// TwinCAT 3 PLC project xpp_pulsepicker_motion
// ProgramVersion: 3.1.4026.17
// libraries:
//   LCLS_MotionAbstraction, * (SLAC)
//   LCLS_Tc_DevAbs, * (SLAC - LCLS)
//   LCLS_Tc_MotSync, * (SLAC - LCLS)
//   Tc2_EtherCAT, * (Beckhoff Automation GmbH)
//   Tc2_MC2, * (Beckhoff Automation GmbH)
//   Tc2_Standard, * (Beckhoff Automation GmbH)
//   Tc2_System, * (Beckhoff Automation GmbH)
//   TcUnit, * (www.tcunit.org)
// project tree:
//   DUTs/ E_HomeIndexState.TcDUT, E_HomeCenterState.TcDUT, E_ModeSelector.TcDUT, E_PickerState.TcDUT, E_PPStatus.TcDUT, E_StatusIndicator.TcDUT, E_ValidationStep.TcDUT, ST_SpeedProfile.TcDUT
//   GVLs/ GVL_Axes.TcGVL, GVL_Common.TcGVL
//   POUs/ FB_FastClose.TcPOU, FB_FastOpen.TcPOU, FB_HomeToCenter.TcPOU, FB_SpindleHomeToCenter.TcPOU, FB_MoveToNearestClosed.TcPOU, FB_PPEPS.TcPOU, FB_SpindleTaskMonitoring.TcPOU, FB_TriggerManagerEL1124.TcPOU (excluded from build), FB_TriggerSetpointManager.TcPOU, PRG_S.TcPOU, PRG_XY.TcPOU
//   POUs/Test/ FB_HomeToCenter_Tests.TcPOU, FB_PPEPS_Tests.TcPOU, PRG_TEST.TcPOU
//   / TestTask.TcTTO, XYTask.TcTTO, STask.TcTTO
// real-time tasks:
//   TASK XYTask: cycle T#5ms, priority 14, ADS port 350
//   TASK STask: cycle T#250us, priority 12, ADS port 351
//   TASK TestTask: cycle T#10ms, priority 16, ADS port 352
// motion (NC):
//   TASK NC-Task 1 SAF: cycle T#250us, priority 4, ADS port 501
//   TASK NC-Task 1 SVB: cycle T#1ms, priority 8, ADS port 511
//   AXIS Y_Test (id 5)
//     OtherSettings: AllowMotionCmdToSlave=true
//     encoder EncType=1
//     drive DrvType=5
//       Analog: TorqueSetpointScale=10, ScaleFactorActTorque=0.1
//       TimeComp: TaskDelayCycles=1
//     controller CtrType=1
//       CtrPara: PriorControlFactor=1
//         Observer: BandWidth=20
//   AXIS X_Test (id 4)
//     OtherSettings: AllowMotionCmdToSlave=true
//     encoder EncType=1
//     drive DrvType=5
//       Analog: TorqueSetpointScale=10, ScaleFactorActTorque=0.1
//       TimeComp: TaskDelayCycles=1
//     controller CtrType=1
//       CtrPara: PriorControlFactor=1
//         Observer: BandWidth=20
//   AXIS Axis_HomeToCenter_Test1 (id 6)
//     OtherSettings: AllowMotionCmdToSlave=true
//     encoder EncType=1
//     drive DrvType=5
//       Analog: TorqueSetpointScale=10, ScaleFactorActTorque=0.1
//     controller CtrType=1
//       CtrPara: PriorControlFactor=1
//         Observer: BandWidth=20
//   AXIS Axis_HomeToCenter_Test2 (id 7)
//     OtherSettings: AllowMotionCmdToSlave=true
//     encoder EncType=1
//     drive DrvType=5
//       Analog: TorqueSetpointScale=10, ScaleFactorActTorque=0.1
//     controller CtrType=1
//       CtrPara: PriorControlFactor=1
//         Observer: BandWidth=20
//   AXIS Axis_HomeToCenter_Test3 (id 8)
//     OtherSettings: AllowMotionCmdToSlave=true
//     encoder EncType=1
//     drive DrvType=5
//       Analog: TorqueSetpointScale=10, ScaleFactorActTorque=0.1
//     controller CtrType=1
//       CtrPara: PriorControlFactor=1
//         Observer: BandWidth=20
//   AXIS Axis_HomeToCenter_Test4 (id 9)
//     OtherSettings: AllowMotionCmdToSlave=true
//     encoder EncType=1
//     drive DrvType=5
//       Analog: TorqueSetpointScale=10, ScaleFactorActTorque=0.1
//     controller CtrType=1
//       CtrPara: PriorControlFactor=1
//         Observer: BandWidth=20
//   AXIS Axis_HomeToCenter_Test5 (id 10)
//     OtherSettings: AllowMotionCmdToSlave=true
//     encoder EncType=1
//     drive DrvType=5
//       Analog: TorqueSetpointScale=10, ScaleFactorActTorque=0.1
//     controller CtrType=1
//       CtrPara: PriorControlFactor=1
//         Observer: BandWidth=20
//   AXIS Y (id 3)
//     Dynamic: AccelerationMaximum=200, DecelerationMaximum=200, Acceleration=134.468, Deceleration=134.468, Jerk=488.416
//     Velo: RefSearch=0.6383, RefSync=0.6383, SlowManual=0.25, FastManual=0.35, Fast=63.83, Maximum=63.83
//     PositionAreaControl: Range=0.1
//     TargetPosControl: Range=0.1
//     PEHControl: Time=1
//     OtherSettings: PulseDistancePos=0.1, PulseDistanceNeg=0.1
//     encoder EncType=19
//       EncPara: ScaleFactorNumerator=5, ScaleFactorDenominator=1048576, EncMode=3, MaxCount=#xffffffff
//         TimeComp: TimeCompMode=1, EncDelayCycles=4
//     drive DrvType=16
//       DrvPara: MaxCount=#xffffffff, DriveControlDWord=#x00020100
//         Analog: VeloReferenz=70.213, VeloScale=32, TorqueSetpointScale=10, ScaleFactorActTorque=0.1
//         TimeComp: TaskDelayCycles=1
//     controller CtrType=2
//       CtrPara: PriorControlFactor=1
//         PosDiffControl: Range=0.1
//         PID: PosKp=0
//         Observer: BandWidth=20
//   AXIS X (id 2)
//     Dynamic: AccelerationMaximum=80, DecelerationMaximum=80, Acceleration=57.5064, Deceleration=57.5064, Jerk=743.932
//     Velo: RefSearch=0.45, RefSync=0.25, SlowManual=0.25, FastManual=0.25, Fast=7.056, Maximum=7.056
//     PositionAreaControl: Range=0.1
//     TargetPosControl: Range=0.1
//     PEHControl: Time=1
//     OtherSettings: PulseDistancePos=0.1, PulseDistanceNeg=0.1
//     encoder EncType=19
//       EncPara: ScaleFactorNumerator=0.635, ScaleFactorDenominator=1048576, EncMode=3, MaxCount=#xffffffff
//         TimeComp: TimeCompMode=1, EncDelayCycles=4
//     drive DrvType=16
//       DrvPara: MaxCount=#xffffffff, DriveControlDWord=#x00020100
//         Analog: VeloReferenz=7.7616, VeloScale=32, TorqueSetpointScale=10, ScaleFactorActTorque=0.1
//         TimeComp: TaskDelayCycles=1
//     controller CtrType=1
//       CtrPara: PriorControlFactor=1
//         PosDiffControl: Range=0.1
//         PID: PosKp=0
//         Observer: BandWidth=20
//   AXIS Spindle (id 1)
//     General: UnitName=°
//     Dynamic: AccelerationMaximum=47150500, DecelerationMaximum=47150500, Acceleration=2512000, Deceleration=2512000, Jerk=2673789830.50848
//     Velo: RefSearch=82.10526, RefSync=82.10526, SlowManual=15.5263, FastManual=25.1578, Fast=14210.526, Maximum=4000
//     PositionAreaControl: Range=0.1
//     TargetPosControl: Range=0.1
//     BacklashCompensation: Range=-1.25
//     OtherSettings: AllowMotionCmdToSlave=true, PulseDistancePos=0.1, PulseDistanceNeg=0.1
//     encoder EncType=19
//       EncPara: ScaleFactorNumerator=360, ScaleFactorDenominator=1048576, MaxCount=#xffffffff
//     drive DrvType=16
//       DrvPara: MaxCount=#xffffffff, DriveControlDWord=#x00020100
//         Analog: VeloReferenz=7200, TorqueSetpointScale=10, ScaleFactorActTorque=0.1
//         TimeComp: TaskDelayCycles=1
//     controller CtrType=2
//       CtrPara: PriorControlFactor=1
//         PosDiffControl: Range=3
//         PID: PosKp=0
//         Observer: BandWidth=20
// I/O:
//   DEVICE Device 1 (EtherCAT), AmsNetId 172.21.86.248.2.1
//     Term 1 (EK1200) [EK1200-5000 EtherCAT Power supply (2A E-Bus)]
//       Dongle [EL6070 1Ch. Licensing-Terminal]
//       Spindle [EL7062-0000 2Ch. Stepper motor output stage (48V, 3A)]
//         startup 28688:3 := 08 // DRV Outputs Ch.1 / Modes of operation
//         startup 28688:16 := FF7F // DRV Outputs Ch.1 / Positive torque limit value
//         startup 28688:17 := FF7F // DRV Outputs Ch.1 / Negative torque limit value
//         startup 32784:87 := 64 // DRV Amplifier Settings Ch.1 / Position loop velocity feed forward gain
//         startup 32784:109 := 64000000 // DRV Amplifier Settings Ch.1 / Torque feed forward gain
//         startup 32785:52 := A00F0000 // DRV Motor Settings Ch.1 / Configured motor current
//         startup 32784:19 := 1A00 // DRV Amplifier Settings Ch.1 / Current loop proportional gain
//         startup 32784:18 := 1300 // DRV Amplifier Settings Ch.1 / Current loop integral time
//         startup 32784:21 := 51000000 // DRV Amplifier Settings Ch.1 / Velocity loop proportional gain
//         startup 32784:20 := 96000000 // DRV Amplifier Settings Ch.1 / Velocity loop integral time
//       XY [EL7062-0000 2Ch. Stepper motor output stage (48V, 3A)]
//         startup 28688:3 := 08 // DRV Outputs Ch.1 / Modes of operation
//         startup 28688:16 := FF7F // DRV Outputs Ch.1 / Positive torque limit value
//         startup 28688:17 := FF7F // DRV Outputs Ch.1 / Negative torque limit value
//         startup 32784:87 := 64 // DRV Amplifier Settings Ch.1 / Position loop velocity feed forward gain
//         startup 32784:109 := 64000000 // DRV Amplifier Settings Ch.1 / Torque feed forward gain
//         startup 32785:52 := C4090000 // DRV Motor Settings Ch.1 / Configured motor current
//         startup 32784:19 := 2800 // DRV Amplifier Settings Ch.1 / Current loop proportional gain
//         startup 32784:18 := 1200 // DRV Amplifier Settings Ch.1 / Current loop integral time
//         startup 32784:21 := 2B000000 // DRV Amplifier Settings Ch.1 / Velocity loop proportional gain
//         startup 32784:20 := 96000000 // DRV Amplifier Settings Ch.1 / Velocity loop integral time
//         startup 33042:19 := 0000 // DRV Brake Settings Ch.2 / Emergency application timeout
//         startup 33040:51 := 0A00 // DRV Amplifier Settings Ch.2 / Stand still window
//         startup 28944:3 := 08 // DRV Outputs Ch.2 / Modes of operation
//         startup 28944:16 := FF7F // DRV Outputs Ch.2 / Positive torque limit value
//         startup 28944:17 := FF7F // DRV Outputs Ch.2 / Negative torque limit value
//         startup 33040:87 := 64 // DRV Amplifier Settings Ch.2 / Position loop velocity feed forward gain
//         startup 33040:109 := 64000000 // DRV Amplifier Settings Ch.2 / Torque feed forward gain
//         startup 33041:52 := A00F0000 // DRV Motor Settings Ch.2 / Configured motor current
//         startup 33040:19 := 3000 // DRV Amplifier Settings Ch.2 / Current loop proportional gain
//         startup 33040:18 := 2700 // DRV Amplifier Settings Ch.2 / Current loop integral time
//         startup 33040:21 := 66000000 // DRV Amplifier Settings Ch.2 / Velocity loop proportional gain
//         startup 33040:20 := 96000000 // DRV Amplifier Settings Ch.2 / Velocity loop integral time
//       Term 5 (EL9505) [EL9505 Power supply terminal 5V]
//       Trigger [EL1124 4Ch. Dig. Input 5V, 10µs, Sensor Power]
//       Term 7 (EL9011) [EL9011 End Terminal]
// variable links:
//   (this object) <-> Device 1 (EtherCAT)/Term 1 (EK1200)/XY
//     Drive/Inputs/In/nDataIn1 <-> DRV Following error actual value Channel 2/Following error actual value
//     Drive/Inputs/In/nDataIn1 <-> DRV Following error actual value Channel 1/Following error actual value
//     Drive/Inputs/In/nDataIn3[0] <-> DRV Torque actual value Channel 2/Torque actual value
//     Drive/Inputs/In/nDataIn3[0] <-> DRV Torque actual value Channel 1/Torque actual value
//     Drive/Inputs/In/nDcOutputTime <-> InfoData/DcOutputShift
//     Drive/Inputs/In/nState1 <-> DRV Statusword Channel 2/Statusword
//     Drive/Inputs/In/nState1 <-> DRV Statusword Channel 1/Statusword
//     Drive/Inputs/In/nState2 <-> DRV Statusword Channel 2/Statusword @bit 8
//     Drive/Inputs/In/nState2 <-> DRV Statusword Channel 1/Statusword @bit 8
//     Drive/Inputs/In/nState4 @bit 1 <-> WcState/InputToggle
//     Drive/Inputs/In/nState4 <-> WcState/WcState
//     Drive/Outputs/Out/nCtrl1 <-> DRV Controlword Channel 2/Controlword
//     Drive/Outputs/Out/nCtrl1 <-> DRV Controlword Channel 1/Controlword
//     Drive/Outputs/Out/nCtrl2 <-> DRV Controlword Channel 2/Controlword @bit 8
//     Drive/Outputs/Out/nCtrl2 <-> DRV Controlword Channel 1/Controlword @bit 8
//     Drive/Outputs/Out/nDataOut1 <-> DRV Target position Channel 2/Target position
//     Drive/Outputs/Out/nDataOut1 <-> DRV Target position Channel 1/Target position
//     Enc/Inputs/In/nDataIn1 <-> FB Position Channel 2/Position
//     Enc/Inputs/In/nDataIn1 <-> FB Position Channel 1/Position
//     Enc/Inputs/In/nDcInputTime <-> InfoData/DcInputShift
//     Enc/Inputs/In/nState4 @bit 1 <-> WcState/InputToggle
//     Enc/Inputs/In/nState4 <-> WcState/WcState
//     XYTask Inputs/PRG_XY.fbX.fbEncoderScaling.nRawEncoderUDINT <-> FB Position Channel 1/Position
//     XYTask Inputs/PRG_XY.fbX.fbLimSwStatus.bLimitBwd <-> DI Inputs Channel 1/Input 1
//     XYTask Inputs/PRG_XY.fbX.fbLimSwStatus.bLimitFwd <-> DI Inputs Channel 1/Input 2
//     XYTask Inputs/PRG_XY.fbY.fbEncoderScaling.nRawEncoderUDINT <-> FB Position Channel 2/Position
//     XYTask Inputs/PRG_XY.fbY.fbLimSwStatus.bLimitBwd <-> DI Inputs Channel 2/Input 2
//     XYTask Inputs/PRG_XY.fbY.fbLimSwStatus.bLimitFwd <-> DI Inputs Channel 2/Input 1
//   (this object) <-> Device 1 (EtherCAT)/Term 1 (EK1200)/Spindle
//     Drive/Inputs/In/nDataIn1 <-> DRV Following error actual value Channel 1/Following error actual value
//     Drive/Inputs/In/nDataIn3[0] <-> DRV Torque actual value Channel 1/Torque actual value
//     Drive/Inputs/In/nState1 <-> DRV Statusword Channel 1/Statusword
//     Drive/Inputs/In/nState2 <-> DRV Statusword Channel 1/Statusword @bit 8
//     Drive/Inputs/In/nState4 @bit 1 <-> WcState/InputToggle
//     Drive/Inputs/In/nState4 <-> WcState/WcState
//     Drive/Outputs/Out/nCtrl1 <-> DRV Controlword Channel 1/Controlword
//     Drive/Outputs/Out/nCtrl2 <-> DRV Controlword Channel 1/Controlword @bit 8
//     Drive/Outputs/Out/nDataOut1 <-> DRV Target position Channel 1/Target position
//     Enc/Inputs/In/nDataIn1 <-> FB Position Channel 1/Position
//     Enc/Inputs/In/nDataIn3 <-> FB Touch probe 1 pos position Channel 1/TP1 Pos position
//     Enc/Inputs/In/nDataIn5 <-> FB Touch probe 2 pos position Channel 1/TP2 Pos position
//     Enc/Inputs/In/nState4 @bit 1 <-> WcState/InputToggle
//     Enc/Inputs/In/nState4 <-> WcState/WcState
//     Enc/Inputs/In/nState5 <-> FB Touch probe status Channel 1/Touch probe status/TP1 Enable
//     Enc/Inputs/In/nState6 <-> FB Touch probe status Channel 1/Touch probe status/TP2 Enable
//     Enc/Inputs/In/nState5 @bit 7 <-> FB Touch probe status Channel 1/Touch probe status/TP1 Input
//     Enc/Inputs/In/nState6 @bit 7 <-> FB Touch probe status Channel 1/Touch probe status/TP2 Input
//     Enc/Inputs/In/nState5 @bit 2 <-> FB Touch probe status Channel 1/Touch probe status/TP1 Neg value stored
//     Enc/Inputs/In/nState6 @bit 2 <-> FB Touch probe status Channel 1/Touch probe status/TP2 Neg value stored
//     Enc/Inputs/In/nState5 @bit 1 <-> FB Touch probe status Channel 1/Touch probe status/TP1 Pos value stored
//     Enc/Inputs/In/nState6 @bit 1 <-> FB Touch probe status Channel 1/Touch probe status/TP2 Pos value stored
//     Enc/Outputs/Out/nCtrl5 @bit 1 <-> FB Touch probe control Channel 1/Touch probe function/TP1 Continous
//     Enc/Outputs/Out/nCtrl6 @bit 1 <-> FB Touch probe control Channel 1/Touch probe function/TP2 Continous
//     Enc/Outputs/Out/nCtrl5 <-> FB Touch probe control Channel 1/Touch probe function/TP1 Enable
//     Enc/Outputs/Out/nCtrl6 <-> FB Touch probe control Channel 1/Touch probe function/TP2 Enable
//     Enc/Outputs/Out/nCtrl5 @bit 5 <-> FB Touch probe control Channel 1/Touch probe function/TP1 Enable neg edge
//     Enc/Outputs/Out/nCtrl6 @bit 5 <-> FB Touch probe control Channel 1/Touch probe function/TP2 Enable neg edge
//     Enc/Outputs/Out/nCtrl5 @bit 4 <-> FB Touch probe control Channel 1/Touch probe function/TP1 Enable pos edge
//     Enc/Outputs/Out/nCtrl6 @bit 4 <-> FB Touch probe control Channel 1/Touch probe function/TP2 Enable pos edge
//     Enc/Outputs/Out/nCtrl5 @bit 2 <-> FB Touch probe control Channel 1/Touch probe function/TP1 Trigger mode
//     Enc/Outputs/Out/nCtrl6 @bit 2 <-> FB Touch probe control Channel 1/Touch probe function/TP2 Trigger mode
//     STask Inputs/PRG_S.fbHomeIdx.bHomeIndex <-> DI Inputs Channel 1/Encoder C
//     STask Inputs/PRG_S.fbS.fbEncoderScaling.nRawEncoderUDINT <-> FB Position Channel 1/Position
//   (this object) <-> Device 1 (EtherCAT)/Term 1 (EK1200)/Trigger
//     STask Inputs/PRG_S.fbTrigMgr.fbTrigSrc.bTrigger <-> Channel 1/Input
//   (this object) <-> NC-Task 1 SAF/Axes/Axis_HomeToCenter_Test1
//     TestTask Inputs/PRG_TEST.fb_HomeToCenter_Tests.fbAxisRef[1].NcToPlc <-> Outputs/ToPlc
//     TestTask Outputs/PRG_TEST.fb_HomeToCenter_Tests.fbAxisRef[1].PlcToNc <-> Inputs/FromPlc
//   (this object) <-> NC-Task 1 SAF/Axes/Axis_HomeToCenter_Test2
//     TestTask Inputs/PRG_TEST.fb_HomeToCenter_Tests.fbAxisRef[2].NcToPlc <-> Outputs/ToPlc
//     TestTask Outputs/PRG_TEST.fb_HomeToCenter_Tests.fbAxisRef[2].PlcToNc <-> Inputs/FromPlc
//   (this object) <-> NC-Task 1 SAF/Axes/Axis_HomeToCenter_Test3
//     TestTask Inputs/PRG_TEST.fb_HomeToCenter_Tests.fbAxisRef[3].NcToPlc <-> Outputs/ToPlc
//     TestTask Outputs/PRG_TEST.fb_HomeToCenter_Tests.fbAxisRef[3].PlcToNc <-> Inputs/FromPlc
//   (this object) <-> NC-Task 1 SAF/Axes/Axis_HomeToCenter_Test4
//     TestTask Inputs/PRG_TEST.fb_HomeToCenter_Tests.fbAxisRef[4].NcToPlc <-> Outputs/ToPlc
//     TestTask Outputs/PRG_TEST.fb_HomeToCenter_Tests.fbAxisRef[4].PlcToNc <-> Inputs/FromPlc
//   (this object) <-> NC-Task 1 SAF/Axes/Axis_HomeToCenter_Test5
//     TestTask Inputs/PRG_TEST.fb_HomeToCenter_Tests.fbAxisRef[5].NcToPlc <-> Outputs/ToPlc
//     TestTask Outputs/PRG_TEST.fb_HomeToCenter_Tests.fbAxisRef[5].PlcToNc <-> Inputs/FromPlc
//   (this object) <-> NC-Task 1 SAF/Axes/Spindle
//     STask Inputs/GVL_Axes.Axes[1].NcToPlc <-> Outputs/ToPlc
//     STask Outputs/GVL_Axes.Axes[1].PlcToNc <-> Inputs/FromPlc
//   (this object) <-> NC-Task 1 SAF/Axes/X
//     STask Inputs/GVL_Axes.Axes[2].NcToPlc <-> Outputs/ToPlc
//     STask Outputs/GVL_Axes.Axes[2].PlcToNc <-> Inputs/FromPlc
//   (this object) <-> NC-Task 1 SAF/Axes/Y
//     STask Inputs/GVL_Axes.Axes[3].NcToPlc <-> Outputs/ToPlc
//     STask Outputs/GVL_Axes.Axes[3].PlcToNc <-> Inputs/FromPlc

CONFIGURATION xpp_pulsepicker_motion
    RESOURCE PLC ON TwinCAT3
        TASK TestTask(INTERVAL := T#10ms, PRIORITY := 16);
        TASK XYTask(INTERVAL := T#5ms, PRIORITY := 14);
        TASK STask(INTERVAL := T#250us, PRIORITY := 12);
        PROGRAM PRG_TEST WITH TestTask : PRG_TEST;
        PROGRAM PRG_XY WITH XYTask : PRG_XY;
        PROGRAM PRG_S WITH STask : PRG_S;
    END_RESOURCE
END_CONFIGURATION

// ---- DUTs/E_HomeIndexState.TcDUT
{attribute 'qualified_only'}
{attribute 'strict'}
{attribute 'to_string'}
TYPE E_HomeIndexState :
(
    Idle := 0,
    Homing,
    WaitHomed,
    HomingUnlatch,
    HomingPulsed,
    WaitHomeDone,
    CenterMove,
    WaitCenterDone,
    SetPosition,
    HomingDone,
    Done,
    Error
)UINT;
END_TYPE

// ---- DUTs/E_HomeCenterState.TcDUT
{attribute 'qualified_only'}
{attribute 'strict'}
{attribute 'to_string'}
TYPE E_HomeCenterState :
(
    Idle           := 0,   // waiting for NC rising edge of bHoming
    WaitHomeDone   := 1,   // drive homing to switch; wait for bDone AND bHomed
    CenterMove     := 2,   // centering AbsoluteMove issued; wait for completion
    WaitCenterDone := 3,   // MC_SetPosition executing to zero the centered position
    HomingDone     := 4,   // restore motion params, return to Idle
    Error          := 5    // latched error; requires Reset()
);
END_TYPE

// ---- DUTs/E_ModeSelector.TcDUT
{attribute 'qualified_only'}
{attribute 'to_string'}
TYPE E_ModeSelector :
(
    ModeNone := 0,
    FlipFlop := 1,
    Burst := 2,
    Open := 3,
    Close := 4,
    Home := 5
) UINT;
END_TYPE

// ---- DUTs/E_PickerState.TcDUT
{attribute 'qualified_only'}
{attribute 'strict'}
{attribute 'to_string'}
TYPE E_PickerState :
(
    Init,           // Startup: Read ModeSelect/SlitStatusFlag from NV
    Ready,
    ModeSelect,     // Idle/waiting for user/command mode selection
    ModeExecute,    // Executing selected mode (One-Shot, Flip-Flop, etc)
    ErrorState      // Error or drift handling and recovery
);
END_TYPE

// ---- DUTs/E_PPStatus.TcDUT
{attribute 'qualified_only'}
{attribute 'strict'}
{attribute 'to_string'}
TYPE E_PPStatus :
(
    UNKNOWN:= 0,
    IN := 1,
    OUT := 2
) UINT;
END_TYPE

// ---- DUTs/E_StatusIndicator.TcDUT
{attribute 'qualified_only'}
{attribute 'strict'}
{attribute 'to_string'}
TYPE E_StatusIndicator :
(
    Init := 10,
    Wait := 11,
    Complete := 12,
    Closed := 13,
    Opened := 14,
    Done := 15,
    // Special states
    HardReset := 80,
    SoftReset := 81
);
END_TYPE

// ---- DUTs/E_ValidationStep.TcDUT
{attribute 'qualified_only'}
{attribute 'strict'}
{attribute 'to_string'}
TYPE E_ValidationStep :
(
    INITIALIZE := 0,
    WAIT_FOR_IDLE,
    COMMAND_SEQUENCE_START,
    GENERATE_TARGET_POINTS,
    COMMAND_MOVE_TO_FIRST_TARGET,
    COMMAND_START_TRIGGERS,
    COMMAND_REVERSE_INT,
    CONFIRM_BACK_TO_IDLE
);
END_TYPE

// ---- DUTs/ST_SpeedProfile.TcDUT
TYPE ST_SpeedProfile :
STRUCT
    InitialVelocity : LREAL;
    MaxVelocity : LREAL;
    Acceleration : LREAL;
    Deceleration : LREAL;
END_STRUCT
END_TYPE

// ---- GVLs/GVL_Axes.TcGVL
{attribute 'qualified_only'}
VAR_GLOBAL
    Axes :  ARRAY[1..4] OF AXIS_REF;
END_VAR

// ---- GVLs/GVL_Common.TcGVL
{attribute 'qualified_only'}
VAR_GLOBAL
    fbPersistentDataStorage : LCLS_Tc_DevAbs.FB_PersistentDataStorage;
    eModeSelect : E_ModeSelector := E_ModeSelector.ModeNone;
END_VAR

// ---- POUs/Test/PRG_TEST.TcPOU
PROGRAM PRG_TEST
VAR
    fb_PPEPS_Tests : FB_PPEPS_Tests;
    {attribute 'TcNcAxis' := '
        .fbAxisRef[1] := Axis_HomeToCenter_Test1;
        .fbAxisRef[2] := Axis_HomeToCenter_Test2;
        .fbAxisRef[3] := Axis_HomeToCenter_Test3;
        .fbAxisRef[4] := Axis_HomeToCenter_Test4;
        .fbAxisRef[5] := Axis_HomeToCenter_Test5;
    '}
    fb_HomeToCenter_Tests : FB_HomeToCenter_Tests;
END_VAR

TcUnit.Run();

END_PROGRAM

// ---- POUs/Test/FB_PPEPS_Tests.TcPOU
FUNCTION_BLOCK FB_PPEPS_Tests EXTENDS FB_TestSuite
VAR
    afbDoubleX : ARRAY[1..19] OF FB_MotionStageNC_TestDouble;
    afbDoubleY : ARRAY[1..19] OF FB_MotionStageNC_TestDouble;
    afbXEPS    : ARRAY[1..19] OF LCLS_MotionAbstraction.FB_EPS;
    afbYEPS    : ARRAY[1..19] OF LCLS_MotionAbstraction.FB_EPS;
END_VAR

// Move-interlock logic
Test_XInCenter_WhenXWithinWindow();
Test_XNotInCenter_WhenXOutsideWindow();
Test_YAboveMed_WhenYExceedsThreshold();
Test_XMoveAllowed_WhenYLow_AndXInRange();
Test_XMoveBlocked_WhenYHigh_AndXOutsideCenter_MovingAway();
Test_XRecovery_WhenYHigh_AndXMovingTowardCenter();
Test_YMoveAllowed_WhenYLow_AndXInCenter();
Test_YMoveBlocked_WhenYHigh_AndXOutsideCenter();

// Homing gates POWER only (directional stays honest)
Test_XHomeAllowed_GatesPower_WhenYBelowMedium();
Test_XHome_YHigh_PowerNotReleased();
Test_YHomeAllowed_GatesPower_WhenXInCenter();
Test_YHome_PickerActive_AllCleared();
Test_Homing_DoesNotForceDirectional_AntiFakeLimit();
Test_XHoming_CommandHeld_NoExecute_NoPower();

// Picker
Test_PickerActive_BlocksXAndY();
Test_PickerIdle_ReleasesEPS();

// Per-axis bypass
Test_XBypass_OverridesBlockedMove();
Test_Bypass_CannotOverridePickerActive();
Test_XBypass_DoesNotReleasePower();

(* Helper: test whether bit nBit is set in nFlags. Retained for fine-grained
   diagnostics; the primary interlock signal asserted by tests is bEPS_OK
   (the per-channel AND-reduction that feeds the drive power/enable interlock). *)
METHOD PRIVATE GetBit : BOOL
VAR_INPUT
    nFlags : UDINT;
    nBit   : INT;
END_VAR
GetBit := (nFlags AND SHL(UDINT#1, nBit)) <> 0;
END_METHOD

// X at 0.0 (inside center window) -> bXInCenter TRUE. Picker idle, move in window.
// Directional forward/backward bEPS_OK TRUE.
METHOD PRIVATE Test_XInCenter_WhenXWithinWindow
VAR_INST
    fbUUT : FB_PPEPS(iXEPS := afbXEPS[1], iYEPS := afbYEPS[1],
                     iXMotionStage := afbDoubleX[1], iYMotionStage := afbDoubleY[1]);
END_VAR
TEST('Test_XInCenter_WhenXWithinWindow');

afbDoubleX[1].MotionStatus.fActPosition := 0.0;
afbDoubleX[1].MotionCmd.fPosition := 0.0;
afbDoubleY[1].MotionStatus.fActPosition := 0.0;

afbDoubleX[1]();
afbDoubleY[1]();
fbUUT(bPickActive := FALSE);

AssertTrue(fbUUT.bXInCenter,
    'bXInCenter should be TRUE when X=0.0');
AssertTrue(afbXEPS[1].EPSForwardEnable.bEPS_OK,
    'X forward bEPS_OK should be TRUE (picker idle, move in window)');
AssertTrue(afbXEPS[1].EPSBackwardEnable.bEPS_OK,
    'X backward bEPS_OK should be TRUE');

TEST_FINISHED();
END_METHOD

// X at 3.0 (outside center) -> bXInCenter FALSE. Y low, full X range, cmd in range
// -> directional forward bEPS_OK TRUE.
METHOD PRIVATE Test_XNotInCenter_WhenXOutsideWindow
VAR_INST
    fbUUT : FB_PPEPS(iXEPS := afbXEPS[2], iYEPS := afbYEPS[2],
                     iXMotionStage := afbDoubleX[2], iYMotionStage := afbDoubleY[2]);
END_VAR
TEST('Test_XNotInCenter_WhenXOutsideWindow');

afbDoubleX[2].MotionStatus.fActPosition := 3.0;
afbDoubleX[2].MotionCmd.fPosition := 3.0;
afbDoubleY[2].MotionStatus.fActPosition := 0.0;

afbDoubleX[2]();
afbDoubleY[2]();
fbUUT(bPickActive := FALSE);

AssertFalse(fbUUT.bXInCenter,
    'bXInCenter should be FALSE when X=3.0');
AssertTrue(afbXEPS[2].EPSForwardEnable.bEPS_OK,
    'X forward bEPS_OK should be TRUE (Y low, full range, cmd in range)');

TEST_FINISHED();
END_METHOD

// Y at 15.0 (above medium) -> bYAboveMed TRUE. X in center so Y move allowed
// -> Y forward bEPS_OK TRUE.
METHOD PRIVATE Test_YAboveMed_WhenYExceedsThreshold
VAR_INST
    fbUUT : FB_PPEPS(iXEPS := afbXEPS[3], iYEPS := afbYEPS[3],
                     iXMotionStage := afbDoubleX[3], iYMotionStage := afbDoubleY[3]);
END_VAR
TEST('Test_YAboveMed_WhenYExceedsThreshold');

afbDoubleX[3].MotionStatus.fActPosition := 0.0;
afbDoubleY[3].MotionStatus.fActPosition := 15.0;
afbDoubleY[3].MotionCmd.fPosition := 15.0;

afbDoubleX[3]();
afbDoubleY[3]();
fbUUT(bPickActive := FALSE);

AssertTrue(fbUUT.bYAboveMed,
    'bYAboveMed should be TRUE when Y=15.0');
AssertTrue(afbYEPS[3].EPSForwardEnable.bEPS_OK,
    'Y forward bEPS_OK should be TRUE (X in center allows Y move)');

TEST_FINISHED();
END_METHOD

// Y low, X cmd within range -> bXMoveAllowed TRUE; directional forward/backward bEPS_OK TRUE.
METHOD PRIVATE Test_XMoveAllowed_WhenYLow_AndXInRange
VAR_INST
    fbUUT : FB_PPEPS(iXEPS := afbXEPS[4], iYEPS := afbYEPS[4],
                     iXMotionStage := afbDoubleX[4], iYMotionStage := afbDoubleY[4]);
END_VAR
TEST('Test_XMoveAllowed_WhenYLow_AndXInRange');

afbDoubleX[4].MotionStatus.fActPosition := 0.0;
afbDoubleX[4].MotionCmd.fPosition := 3.0;
afbDoubleY[4].MotionStatus.fActPosition := 5.0;

afbDoubleX[4]();
afbDoubleY[4]();
fbUUT(bPickActive := FALSE);

AssertTrue(fbUUT.bXMoveAllowed,
    'bXMoveAllowed should be TRUE when Y low and X cmd=3.0');
AssertTrue(afbXEPS[4].EPSForwardEnable.bEPS_OK,
    'X forward bEPS_OK should be TRUE');
AssertTrue(afbXEPS[4].EPSBackwardEnable.bEPS_OK,
    'X backward bEPS_OK should be TRUE');

TEST_FINISHED();
END_METHOD

// Y high, X outside center, cmd further from center -> bXMoveAllowed FALSE.
// Directional bit1=0 -> forward/backward bEPS_OK FALSE.
METHOD PRIVATE Test_XMoveBlocked_WhenYHigh_AndXOutsideCenter_MovingAway
VAR_INST
    fbUUT : FB_PPEPS(iXEPS := afbXEPS[5], iYEPS := afbYEPS[5],
                     iXMotionStage := afbDoubleX[5], iYMotionStage := afbDoubleY[5]);
END_VAR
TEST('Test_XMoveBlocked_WhenYHigh_AndXOutsideCenter_MovingAway');

afbDoubleX[5].MotionStatus.fActPosition := 3.0;
afbDoubleX[5].MotionCmd.fPosition := 4.0;
afbDoubleY[5].MotionStatus.fActPosition := 15.0;

afbDoubleX[5]();
afbDoubleY[5]();
fbUUT(bPickActive := FALSE);

AssertFalse(fbUUT.bXMoveAllowed,
    'bXMoveAllowed should be FALSE when Y high and X moving away from center');
AssertFalse(afbXEPS[5].EPSForwardEnable.bEPS_OK,
    'X forward bEPS_OK should be FALSE (move bit cleared)');
AssertFalse(afbXEPS[5].EPSBackwardEnable.bEPS_OK,
    'X backward bEPS_OK should be FALSE (move bit cleared)');

TEST_FINISHED();
END_METHOD

// Y high, X outside center, cmd toward center -> recovery allowed.
// bXTowardCenter TRUE, bXMoveAllowed TRUE, forward bEPS_OK TRUE.
METHOD PRIVATE Test_XRecovery_WhenYHigh_AndXMovingTowardCenter
VAR_INST
    fbUUT : FB_PPEPS(iXEPS := afbXEPS[6], iYEPS := afbYEPS[6],
                     iXMotionStage := afbDoubleX[6], iYMotionStage := afbDoubleY[6]);
END_VAR
TEST('Test_XRecovery_WhenYHigh_AndXMovingTowardCenter');

afbDoubleX[6].MotionStatus.fActPosition := 3.0;
afbDoubleX[6].MotionCmd.fPosition := 0.0;
afbDoubleY[6].MotionStatus.fActPosition := 15.0;

afbDoubleX[6]();
afbDoubleY[6]();
fbUUT(bPickActive := FALSE);

AssertTrue(fbUUT.bXTowardCenter,
    'bXTowardCenter should be TRUE');
AssertTrue(fbUUT.bXMoveAllowed,
    'bXMoveAllowed should be TRUE for recovery move toward center');
AssertTrue(afbXEPS[6].EPSForwardEnable.bEPS_OK,
    'X forward bEPS_OK should be TRUE (recovery permitted)');

TEST_FINISHED();
END_METHOD

// Y low, X in center, Y cmd within range -> bYMoveAllowed TRUE.
// Y forward/backward bEPS_OK TRUE.
METHOD PRIVATE Test_YMoveAllowed_WhenYLow_AndXInCenter
VAR_INST
    fbUUT : FB_PPEPS(iXEPS := afbXEPS[7], iYEPS := afbYEPS[7],
                     iXMotionStage := afbDoubleX[7], iYMotionStage := afbDoubleY[7]);
END_VAR
TEST('Test_YMoveAllowed_WhenYLow_AndXInCenter');

afbDoubleX[7].MotionStatus.fActPosition := 0.0;
afbDoubleY[7].MotionStatus.fActPosition := 5.0;
afbDoubleY[7].MotionCmd.fPosition := 18.0;

afbDoubleX[7]();
afbDoubleY[7]();
fbUUT(bPickActive := FALSE);

AssertTrue(fbUUT.bYMoveAllowed,
    'bYMoveAllowed should be TRUE when Y low, X in center, cmd=18.0');
AssertTrue(afbYEPS[7].EPSForwardEnable.bEPS_OK,
    'Y forward bEPS_OK should be TRUE');
AssertTrue(afbYEPS[7].EPSBackwardEnable.bEPS_OK,
    'Y backward bEPS_OK should be TRUE');

TEST_FINISHED();
END_METHOD

// Y high, X outside center -> all Y motion blocked. Y forward/backward bEPS_OK FALSE.
METHOD PRIVATE Test_YMoveBlocked_WhenYHigh_AndXOutsideCenter
VAR_INST
    fbUUT : FB_PPEPS(iXEPS := afbXEPS[8], iYEPS := afbYEPS[8],
                     iXMotionStage := afbDoubleX[8], iYMotionStage := afbDoubleY[8]);
END_VAR
TEST('Test_YMoveBlocked_WhenYHigh_AndXOutsideCenter');

afbDoubleX[8].MotionStatus.fActPosition := 3.0;
afbDoubleY[8].MotionStatus.fActPosition := 15.0;
afbDoubleY[8].MotionCmd.fPosition := 5.0;

afbDoubleX[8]();
afbDoubleY[8]();
fbUUT(bPickActive := FALSE);

AssertFalse(fbUUT.bYMoveAllowed,
    'bYMoveAllowed should be FALSE when Y high and X outside center');
AssertFalse(afbYEPS[8].EPSForwardEnable.bEPS_OK,
    'Y forward bEPS_OK should be FALSE');
AssertFalse(afbYEPS[8].EPSBackwardEnable.bEPS_OK,
    'Y backward bEPS_OK should be FALSE');

TEST_FINISHED();
END_METHOD

// Fresh HOME on X with Y below medium -> X-homing ALLOWED. Homing gates POWER only:
// power bEPS_OK TRUE (bXHomeAllowed releases power bit1). Directional follows the
// real move interlock (cmd=0.0 in range, Y low) -> forward bEPS_OK TRUE independently.
METHOD PRIVATE Test_XHomeAllowed_GatesPower_WhenYBelowMedium
VAR_INST
    fbUUT : FB_PPEPS(iXEPS := afbXEPS[9], iYEPS := afbYEPS[9],
                     iXMotionStage := afbDoubleX[9], iYMotionStage := afbDoubleY[9]);
END_VAR
TEST('Test_XHomeAllowed_GatesPower_WhenYBelowMedium');

afbDoubleX[9].MotionStatus.fActPosition := 3.0;
afbDoubleX[9].MotionCmd.fPosition := 0.0;
afbDoubleX[9].MotionStatus.eCommand := E_EpicsMotorCmd.HOME;
afbDoubleX[9].ExMotionStatus.bExecute := TRUE;
afbDoubleY[9].MotionStatus.fActPosition := 5.0;

afbDoubleX[9]();
afbDoubleY[9]();
fbUUT(bPickActive := FALSE);

AssertTrue(fbUUT.bXHoming,
    'bXHoming should be TRUE for fresh HOME request');
AssertTrue(fbUUT.bXHomeAllowed,
    'bXHomeAllowed should be TRUE when Y below medium');
AssertTrue(afbXEPS[9].EPSPowerEnable.bEPS_OK,
    'X power bEPS_OK should be TRUE (homing allowed releases power)');
AssertTrue(afbXEPS[9].EPSForwardEnable.bEPS_OK,
    'X forward bEPS_OK should be TRUE (move interlock allows it; homing does not gate direction)');

TEST_FINISHED();
END_METHOD

// Fresh HOME on X but Y HIGH -> bXHomeAllowed = NOT bYAboveMed = FALSE.
// Homing gates POWER: power bit1 = bXHomeAllowed = FALSE -> X power bEPS_OK FALSE.
// Directional is independent and here also blocked (Y high, cmd away) -> forward bEPS_OK FALSE.
METHOD PRIVATE Test_XHome_YHigh_PowerNotReleased
VAR_INST
    fbUUT : FB_PPEPS(iXEPS := afbXEPS[10], iYEPS := afbYEPS[10],
                     iXMotionStage := afbDoubleX[10], iYMotionStage := afbDoubleY[10]);
END_VAR
TEST('Test_XHome_YHigh_PowerNotReleased');

afbDoubleX[10].MotionStatus.fActPosition := 3.0;
afbDoubleX[10].MotionCmd.fPosition := 4.0;
afbDoubleX[10].MotionStatus.eCommand := E_EpicsMotorCmd.HOME;
afbDoubleX[10].ExMotionStatus.bExecute := TRUE;
afbDoubleY[10].MotionStatus.fActPosition := 15.0;

afbDoubleX[10]();
afbDoubleY[10]();
fbUUT(bPickActive := FALSE);

AssertTrue(fbUUT.bXHoming,
    'bXHoming should be TRUE (request is live)');
AssertFalse(fbUUT.bXHomeAllowed,
    'bXHomeAllowed should be FALSE when Y high');
AssertFalse(afbXEPS[10].EPSPowerEnable.bEPS_OK,
    'X power bEPS_OK should be FALSE (home not allowed gates power)');

TEST_FINISHED();
END_METHOD

// Fresh HOME on Y, X in center, picker idle -> Y-homing ALLOWED. Power bEPS_OK TRUE.
// Directional follows the real move interlock independently.
METHOD PRIVATE Test_YHomeAllowed_GatesPower_WhenXInCenter
VAR_INST
    fbUUT : FB_PPEPS(iXEPS := afbXEPS[11], iYEPS := afbYEPS[11],
                     iXMotionStage := afbDoubleX[11], iYMotionStage := afbDoubleY[11]);
END_VAR
TEST('Test_YHomeAllowed_GatesPower_WhenXInCenter');

afbDoubleX[11].MotionStatus.fActPosition := 0.0;
afbDoubleY[11].MotionStatus.fActPosition := 0.0;
afbDoubleY[11].MotionCmd.fPosition := 0.0;
afbDoubleY[11].MotionStatus.eCommand := E_EpicsMotorCmd.HOME;
afbDoubleY[11].ExMotionStatus.bExecute := TRUE;

afbDoubleX[11]();
afbDoubleY[11]();
fbUUT(bPickActive := FALSE);

AssertTrue(fbUUT.bYHoming,
    'bYHoming should be TRUE for fresh HOME request');
AssertTrue(fbUUT.bYHomeAllowed,
    'bYHomeAllowed should be TRUE when X in center and picker idle');
AssertTrue(afbYEPS[11].EPSPowerEnable.bEPS_OK,
    'Y power bEPS_OK should be TRUE (homing allowed releases power)');

TEST_FINISHED();
END_METHOD

// Fresh HOME on Y, X in center, picker ACTIVE -> picker overrides all.
// bYHomeAllowed forced FALSE; all three Y bEPS_OK FALSE (bit0 held 0 everywhere).
METHOD PRIVATE Test_YHome_PickerActive_AllCleared
VAR_INST
    fbUUT : FB_PPEPS(iXEPS := afbXEPS[12], iYEPS := afbYEPS[12],
                     iXMotionStage := afbDoubleX[12], iYMotionStage := afbDoubleY[12]);
END_VAR
TEST('Test_YHome_PickerActive_AllCleared');

afbDoubleX[12].MotionStatus.fActPosition := 0.0;
afbDoubleY[12].MotionStatus.fActPosition := 0.0;
afbDoubleY[12].MotionStatus.eCommand := E_EpicsMotorCmd.HOME;
afbDoubleY[12].ExMotionStatus.bExecute := TRUE;

afbDoubleX[12]();
afbDoubleY[12]();
fbUUT(bPickActive := TRUE);

AssertFalse(fbUUT.bYHomeAllowed,
    'bYHomeAllowed should be FALSE under picker active');
AssertFalse(afbYEPS[12].EPSPowerEnable.bEPS_OK,
    'Y power bEPS_OK should be FALSE (picker active)');
AssertFalse(afbYEPS[12].EPSForwardEnable.bEPS_OK,
    'Y forward bEPS_OK should be FALSE (picker active)');

TEST_FINISHED();
END_METHOD

// CORE GUARANTEE: during an ALLOWED home, the directional EPS must still follow the
// real move interlock - homing must NOT force the directional bit (which would fake a
// limit switch). Setup: X home allowed (Y low) but a directional move that is blocked.
// Expect: X power bEPS_OK TRUE (home authorized power) AND X forward bEPS_OK FALSE
// (directional honestly blocked). The two channels decouple - that is the design.
METHOD PRIVATE Test_Homing_DoesNotForceDirectional_AntiFakeLimit
VAR_INST
    fbUUT : FB_PPEPS(iXEPS := afbXEPS[13], iYEPS := afbYEPS[13],
                     iXMotionStage := afbDoubleX[13], iYMotionStage := afbDoubleY[13]);
END_VAR
TEST('Test_Homing_DoesNotForceDirectional_AntiFakeLimit');

afbDoubleX[13].MotionStatus.fActPosition := 8.0;   // outside full range so move blocked
afbDoubleX[13].MotionCmd.fPosition := 9.0;          // cmd out of [fXLimMin, fXLimMax]
afbDoubleX[13].MotionStatus.eCommand := E_EpicsMotorCmd.HOME;
afbDoubleX[13].ExMotionStatus.bExecute := TRUE;
afbDoubleY[13].MotionStatus.fActPosition := 5.0;   // below medium -> X-homing allowed

afbDoubleX[13]();
afbDoubleY[13]();
fbUUT(bPickActive := FALSE);

AssertTrue(fbUUT.bXHoming,
    'bXHoming should be TRUE');
AssertTrue(fbUUT.bXHomeAllowed,
    'bXHomeAllowed should be TRUE (Y below medium)');
AssertTrue(afbXEPS[13].EPSPowerEnable.bEPS_OK,
    'X power bEPS_OK should be TRUE (home authorizes power)');
AssertFalse(fbUUT.bXMoveAllowed,
    'bXMoveAllowed should be FALSE (cmd out of range) - homing must not force it');
AssertFalse(afbXEPS[13].EPSForwardEnable.bEPS_OK,
    'X forward bEPS_OK should be FALSE (directional follows real move interlock, not homing)');

TEST_FINISHED();
END_METHOD

// REGRESSION for the latch bug: eCommand stays HOME but bExecute FALSE (stale, held
// selection). bXHoming MUST be FALSE so the power channel is released normally (not
// gated by a phantom home) and the directional channel follows the move interlock.
METHOD PRIVATE Test_XHoming_CommandHeld_NoExecute_NoPower
VAR_INST
    fbUUT : FB_PPEPS(iXEPS := afbXEPS[14], iYEPS := afbYEPS[14],
                     iXMotionStage := afbDoubleX[14], iYMotionStage := afbDoubleY[14]);
END_VAR
TEST('Test_XHoming_CommandHeld_NoExecute_NoPower');

afbDoubleX[14].MotionStatus.fActPosition := 3.0;
afbDoubleX[14].MotionCmd.fPosition := 0.0;             // an allowed move (Y low)
afbDoubleX[14].MotionStatus.eCommand := E_EpicsMotorCmd.HOME; // command still reads HOME...
afbDoubleX[14].ExMotionStatus.bExecute := FALSE;                // ...but no fresh execute
afbDoubleY[14].MotionStatus.fActPosition := 5.0;

afbDoubleX[14]();
afbDoubleY[14]();
fbUUT(bPickActive := FALSE);

AssertFalse(fbUUT.bXHoming,
    'bXHoming should be FALSE when no fresh execute (latch regression)');
AssertTrue(afbXEPS[14].EPSPowerEnable.bEPS_OK,
    'X power bEPS_OK should be TRUE (not homing -> power released normally)');

TEST_FINISHED();
END_METHOD

// Picker active -> all three bEPS_OK FALSE on both axes (bit0 held 0 everywhere).
METHOD PRIVATE Test_PickerActive_BlocksXAndY
VAR_INST
    fbUUT : FB_PPEPS(iXEPS := afbXEPS[15], iYEPS := afbYEPS[15],
                     iXMotionStage := afbDoubleX[15], iYMotionStage := afbDoubleY[15]);
END_VAR
TEST('Test_PickerActive_BlocksXAndY');

afbDoubleX[15].MotionStatus.fActPosition := 0.0;
afbDoubleX[15].MotionCmd.fPosition := 3.0;
afbDoubleY[15].MotionStatus.fActPosition := 5.0;
afbDoubleY[15].MotionCmd.fPosition := 8.0;

afbDoubleX[15]();
afbDoubleY[15]();
fbUUT(bPickActive := TRUE);

AssertFalse(afbXEPS[15].EPSForwardEnable.bEPS_OK,
    'X forward bEPS_OK should be FALSE (picker active)');
AssertFalse(afbXEPS[15].EPSPowerEnable.bEPS_OK,
    'X power bEPS_OK should be FALSE (picker active)');
AssertFalse(afbYEPS[15].EPSForwardEnable.bEPS_OK,
    'Y forward bEPS_OK should be FALSE (picker active)');
AssertFalse(afbYEPS[15].EPSPowerEnable.bEPS_OK,
    'Y power bEPS_OK should be FALSE (picker active)');

TEST_FINISHED();
END_METHOD

// Picker idle with a valid in-range state -> directional forward/backward bEPS_OK TRUE both axes.
METHOD PRIVATE Test_PickerIdle_ReleasesEPS
VAR_INST
    fbUUT : FB_PPEPS(iXEPS := afbXEPS[16], iYEPS := afbYEPS[16],
                     iXMotionStage := afbDoubleX[16], iYMotionStage := afbDoubleY[16]);
END_VAR
TEST('Test_PickerIdle_ReleasesEPS');

afbDoubleX[16].MotionStatus.fActPosition := 0.0;
afbDoubleY[16].MotionStatus.fActPosition := 0.0;

afbDoubleX[16]();
afbDoubleY[16]();
fbUUT(bPickActive := FALSE);

AssertTrue(afbXEPS[16].EPSForwardEnable.bEPS_OK,
    'X forward bEPS_OK should be TRUE when picker idle');
AssertTrue(afbXEPS[16].EPSBackwardEnable.bEPS_OK,
    'X backward bEPS_OK should be TRUE when picker idle');
AssertTrue(afbYEPS[16].EPSForwardEnable.bEPS_OK,
    'Y forward bEPS_OK should be TRUE when picker idle');

TEST_FINISHED();
END_METHOD

// Per-axis bypass forces the DIRECTIONAL move bit TRUE even when the interlock blocks
// (Y high, X outside, cmd away). Picker idle -> X forward/backward bEPS_OK TRUE.
// Y not bypassed and blocked -> Y forward bEPS_OK FALSE.
METHOD PRIVATE Test_XBypass_OverridesBlockedMove
VAR_INST
    fbUUT : FB_PPEPS(iXEPS := afbXEPS[17], iYEPS := afbYEPS[17],
                     iXMotionStage := afbDoubleX[17], iYMotionStage := afbDoubleY[17]);
END_VAR
TEST('Test_XBypass_OverridesBlockedMove');

afbDoubleX[17].MotionStatus.fActPosition := 3.0;
afbDoubleX[17].MotionCmd.fPosition := 4.0;   // normally blocked
afbDoubleY[17].MotionStatus.fActPosition := 15.0;

fbUUT.bXBypass := TRUE;
fbUUT.bYBypass := FALSE;

afbDoubleX[17]();
afbDoubleY[17]();
fbUUT(bPickActive := FALSE);

AssertTrue(afbXEPS[17].EPSForwardEnable.bEPS_OK,
    'X forward bEPS_OK should be TRUE (bypass forces move bit, picker idle)');
AssertTrue(afbXEPS[17].EPSBackwardEnable.bEPS_OK,
    'X backward bEPS_OK should be TRUE (bypass forces move bit)');
AssertFalse(afbYEPS[17].EPSForwardEnable.bEPS_OK,
    'Y forward bEPS_OK should be FALSE (Y not bypassed, move blocked)');

TEST_FINISHED();
END_METHOD

// SAFETY: bypass on BOTH axes must NOT defeat the picker. With picker active, the
// NOT bPickActive wrapper holds directional bit1 = 0 and bit0 = 0 -> all bEPS_OK FALSE.
METHOD PRIVATE Test_Bypass_CannotOverridePickerActive
VAR_INST
    fbUUT : FB_PPEPS(iXEPS := afbXEPS[18], iYEPS := afbYEPS[18],
                     iXMotionStage := afbDoubleX[18], iYMotionStage := afbDoubleY[18]);
END_VAR
TEST('Test_Bypass_CannotOverridePickerActive');

afbDoubleX[18].MotionStatus.fActPosition := 0.0;
afbDoubleX[18].MotionCmd.fPosition := 0.0;
afbDoubleY[18].MotionStatus.fActPosition := 5.0;
afbDoubleY[18].MotionCmd.fPosition := 5.0;

fbUUT.bXBypass := TRUE;
fbUUT.bYBypass := TRUE;

afbDoubleX[18]();
afbDoubleY[18]();
fbUUT(bPickActive := TRUE);

AssertFalse(afbXEPS[18].EPSForwardEnable.bEPS_OK,
    'X forward bEPS_OK must stay FALSE (picker active, bypass cannot override)');
AssertFalse(afbYEPS[18].EPSForwardEnable.bEPS_OK,
    'Y forward bEPS_OK must stay FALSE (picker active, bypass cannot override)');

TEST_FINISHED();
END_METHOD

// Bypass touches the DIRECTIONAL channel only. With X home requested but NOT allowed
// (Y high), bypass forces the directional bit but must NOT release power: power is gated
// by homing, which bypass does not touch -> X power bEPS_OK FALSE while forward bEPS_OK TRUE.
METHOD PRIVATE Test_XBypass_DoesNotReleasePower
VAR_INST
    fbUUT : FB_PPEPS(iXEPS := afbXEPS[19], iYEPS := afbYEPS[19],
                     iXMotionStage := afbDoubleX[19], iYMotionStage := afbDoubleY[19]);
END_VAR
TEST('Test_XBypass_DoesNotReleasePower');

afbDoubleX[19].MotionStatus.fActPosition := 3.0;
afbDoubleX[19].MotionCmd.fPosition := 4.0;
afbDoubleX[19].MotionStatus.eCommand := E_EpicsMotorCmd.HOME;
afbDoubleX[19].ExMotionStatus.bExecute := TRUE;
afbDoubleY[19].MotionStatus.fActPosition := 15.0;   // Y high -> home not allowed

fbUUT.bXBypass := TRUE;

afbDoubleX[19]();
afbDoubleY[19]();
fbUUT(bPickActive := FALSE);

AssertTrue(afbXEPS[19].EPSForwardEnable.bEPS_OK,
    'X forward bEPS_OK should be TRUE (bypass forces directional bit)');
AssertFalse(afbXEPS[19].EPSPowerEnable.bEPS_OK,
    'X power bEPS_OK should be FALSE (bypass does not touch power; home not allowed)');

TEST_FINISHED();
END_METHOD

END_FUNCTION_BLOCK

// ---- POUs/FB_PPEPS.TcPOU
//  Pulse-picker EPS interlock for the X/Y stage.
//
//  EPS channel model: each FB_EPS channel (forward / backward / power) ANDs all
//  its bits into a per-channel bEPS_OK. The drive section enables/powers a
//  channel only when that channel's bEPS_OK is TRUE (every bit released).
//
//  Homing gates the POWER channel ONLY.
FUNCTION_BLOCK FB_PPEPS
VAR_INPUT
    bPickActive : BOOL;
    {attribute 'pytmc' := '
        pv: 02:bXEpsBypass
        io: io
        field: DESC X ByPass EPS
    '}
    bXBypass: BOOL;
    {attribute 'pytmc' := '
        pv: 03:bYEpsBypass
        io: io
        field: DESC Y ByPass EPS
    '}
    bYBypass : BOOL;
END_VAR
VAR
    iXMotionStage	: I_MotionStage;
    iYMotionStage	: I_MotionStage;
    iXEPS : I_EPS;
    iYEPS : I_EPS;
    bXHoming : BOOL;
    bYHoming : BOOL;
    yMin     : LREAL;
    yMax     : LREAL;
END_VAR

VAR_OUTPUT
    bXMoveAllowed  : BOOL;
    bYMoveAllowed  : BOOL;
    bXHomeAllowed  : BOOL;
    bYHomeAllowed  : BOOL;
    bXInCenter     : BOOL;
    bYAboveMed     : BOOL;
    bXTowardCenter : BOOL;
END_VAR

VAR PERSISTENT
    {attribute 'pytmc' := '
        pv: 02:fXLimMin
        io: i
        field: DESC X Travel Limit Min
    '}
    fXLimMin : LREAL := -5.1;

    {attribute 'pytmc' := '
        pv: 02:fXLimMax
        io: i
        field: DESC X Travel Limit Max
    '}
    fXLimMax : LREAL := 5.1;

    {attribute 'pytmc' := '
        pv: 02:fXCenterLimMin
        io: i
        field: DESC X Center Window Min
    '}
    fXCenterLimMin : LREAL := -0.5;

    {attribute 'pytmc' := '
        pv: 02:fXCenterLimMax
        io: i
        field: DESC X Center Window Max
    '}
    fXCenterLimMax : LREAL := 0.5;

    {attribute 'pytmc' := '
        pv: 03:fYLimMin
        io: i
        field: DESC Y Travel Limit Min
    '}
    fYLimMin : LREAL := -0.1;

    {attribute 'pytmc' := '
        pv: 03:fYLimMedium
        io: i
        field: DESC Y Critical Threshold
    '}
    fYLimMedium : LREAL := 10.0;

    {attribute 'pytmc' := '
        pv: 03:fYLimMax
        io: i
        field: DESC Y Travel Limit Max
    '}
    fYLimMax : LREAL := 20.1;
END_VAR

bXInCenter := (iXMotionStage.MotionStatus.fActPosition >= fXCenterLimMin) AND
              (iXMotionStage.MotionStatus.fActPosition <= fXCenterLimMax);
bYAboveMed := iYMotionStage.MotionStatus.fActPosition > fYLimMedium;

//  bExecute is the drive-section confirmation of a FRESH home request; combined
//  with eCommand=HOME it distinguishes a live request from a stale, held command
bXHoming := iXMotionStage.ExMotionStatus.bNewMoveReq AND (iXMotionStage.MotionStatus.eCommand = E_EpicsMotorCmd.HOME);
bYHoming := iYMotionStage.ExMotionStatus.bNewMoveReq AND (iYMotionStage.MotionStatus.eCommand = E_EpicsMotorCmd.HOME);

//  Y move interlock
yMin := fYLimMin;
IF bYAboveMed THEN
    bYMoveAllowed := bXInCenter;
ELSE
    yMax := SEL(bXInCenter, fYLimMedium, fYLimMax);
    bYMoveAllowed := (iYMotionStage.MotionCmd.fPosition >= yMin) AND
                     (iYMotionStage.MotionCmd.fPosition <= yMax);
END_IF

//  X move interlock
IF bYAboveMed THEN
    IF bXInCenter THEN
        bXMoveAllowed := (iXMotionStage.MotionCmd.fPosition >= fXCenterLimMin) AND
                         (iXMotionStage.MotionCmd.fPosition <= fXCenterLimMax);
    ELSE
        //  Outside center with Y high: only allow motion that moves TOWARD center.
        bXTowardCenter := (iXMotionStage.MotionStatus.fActPosition < fXCenterLimMin AND
                           iXMotionStage.MotionCmd.fPosition > iXMotionStage.MotionStatus.fActPosition) OR
                          (iXMotionStage.MotionStatus.fActPosition > fXCenterLimMax AND
                           iXMotionStage.MotionCmd.fPosition < iXMotionStage.MotionStatus.fActPosition);
        bXMoveAllowed := bXTowardCenter;
    END_IF
ELSE
    bXMoveAllowed := (iXMotionStage.MotionCmd.fPosition >= fXLimMin) AND
                     (iXMotionStage.MotionCmd.fPosition <= fXLimMax);
END_IF

//  Y homing interlock: gates POWER only, never directional
IF bYHoming THEN
    bYHomeAllowed := bXInCenter;
ELSE
    bYHomeAllowed := TRUE;
END_IF

//  X homing interlock: gates POWER only, never directional
IF bXHoming THEN
    bXHomeAllowed := NOT bYAboveMed;
ELSE
    bXHomeAllowed := TRUE;
END_IF

//  Picker active overrules all
//  The EPS bit writes below also enforce this at the bit level (picker bit0 and
//  the NOT bPickActive wrapper on the move bit).
IF bPickActive THEN
    bXMoveAllowed := FALSE;
    bYMoveAllowed := FALSE;
    bXHomeAllowed := FALSE;
    bYHomeAllowed := FALSE;
END_IF

//
//  DIRECTIONAL (forward / backward):
//    bit 0 : picker gate  NOT bPickActive, never bypassable
//    bit 1 : move interlock OR bypass, picker still absolute
//            = NOT bPickActive AND (bBypass OR bMoveAllowed)
//    Gated by the MOVE interlock only; NEVER by homing (avoids faking the limit
//    switch). Both bits 1 => directional bEPS_OK TRUE.
//
//  POWER:
//    bit 0 : picker gate  NOT bPickActive, never bypassable
//    bit 1 : homing gate  SEL(bHoming, TRUE, bHomeAllowed)
//            not homing       -> TRUE  (released; power depends only on picker)
//            homing requested -> bHomeAllowed (TRUE only if home permitted)
//    Both bits 1 => power bEPS_OK TRUE => drive section grants power.
//    Bypass does NOT touch the power channel.

//  X directional: move interlock + bypass, picker absolute
iXEPS.setBitForward (nBits := 0, bValue := NOT bPickActive);
iXEPS.setBitBackward(nBits := 0, bValue := NOT bPickActive);
iXEPS.setBitForward (nBits := 1, bValue := NOT bPickActive AND (bXBypass OR bXMoveAllowed));
iXEPS.setBitBackward(nBits := 1, bValue := NOT bPickActive AND (bXBypass OR bXMoveAllowed));
//  X power: picker gate + homing gate (not bypassable)
iXEPS.setBitPower   (nBits := 0, bValue := NOT bPickActive);
iXEPS.setBitPower   (nBits := 1, bValue := SEL(bXHoming, TRUE, bXHomeAllowed));

//  Y directional: move interlock + bypass, picker absolute
iYEPS.setBitForward (nBits := 0, bValue := NOT bPickActive);
iYEPS.setBitBackward(nBits := 0, bValue := NOT bPickActive);
iYEPS.setBitForward (nBits := 1, bValue := NOT bPickActive AND (bYBypass OR bYMoveAllowed));
iYEPS.setBitBackward(nBits := 1, bValue := NOT bPickActive AND (bYBypass OR bYMoveAllowed));
//  Y power - picker gate + homing gate (not bypassable)
iYEPS.setBitPower   (nBits := 0, bValue := NOT bPickActive);
iYEPS.setBitPower   (nBits := 1, bValue := SEL(bYHoming, TRUE, bYHomeAllowed));

//FB_Init is always available implicitly and it is used primarily for initialization.
//The return value is not evaluated. For a specific influence, you can also declare the
//methods explicitly and provide additional code there with the standard initialization
//code. You can evaluate the return value.
METHOD FB_Init: BOOL
VAR_INPUT
    bInitRetains: BOOL; // TRUE: the retain variables are initialized (reset warm / reset cold)
    bInCopyCode: BOOL;  // TRUE: the instance will be copied to the copy code afterward (online change)
    iXMotionStage	: I_MotionStage;
    iYMotionStage	: I_MotionStage;
    iXEPS : I_EPS;
    iYEPS : I_EPS;
END_VAR
THIS^.iXMotionStage := iXMotionStage;
THIS^.iYMotionStage := iYMotionStage;
THIS^.iXEPS := iXEPS;
THIS^.iYEPS := iYEPS;
END_METHOD

END_FUNCTION_BLOCK

// ---- POUs/Test/FB_HomeToCenter_Tests.TcPOU
FUNCTION_BLOCK FB_HomeToCenter_Tests EXTENDS FB_TestSuite
VAR
    //  Real stages + axes + persistent-storage doubles (one per test pair).
    fbAxisRef               : ARRAY[1..5] OF AXIS_REF;
    fbPersistentDataStorage : ARRAY[1..5] OF LCLS_Tc_DevAbs.FB_PersistentDataStorageTestDouble;
    afbStage : ARRAY[1..5] OF FB_MotionStageNC[
        (sName := 'HC_T1', AxisRef := fbAxisRef[1], iPersistentDataStorage := fbPersistentDataStorage[1]),
        (sName := 'HC_T2', AxisRef := fbAxisRef[2], iPersistentDataStorage := fbPersistentDataStorage[2]),
        (sName := 'HC_T3', AxisRef := fbAxisRef[3], iPersistentDataStorage := fbPersistentDataStorage[3]),
        (sName := 'HC_T4', AxisRef := fbAxisRef[4], iPersistentDataStorage := fbPersistentDataStorage[4]),
        (sName := 'HC_T5', AxisRef := fbAxisRef[5], iPersistentDataStorage := fbPersistentDataStorage[5])
    ] := [
        (RestoreMotionParams := FALSE, DoNotRestoreNcParameters := TRUE),
        (RestoreMotionParams := FALSE, DoNotRestoreNcParameters := TRUE),
        (RestoreMotionParams := FALSE, DoNotRestoreNcParameters := TRUE),
        (RestoreMotionParams := FALSE, DoNotRestoreNcParameters := TRUE),
        (RestoreMotionParams := FALSE, DoNotRestoreNcParameters := TRUE)
    ];
    bStagesInit : BOOL := TRUE;
    nInit       : INT;
END_VAR

// One-time mode/limit enable for all stages (mirrors the T10 first-scan block).
// HomeEnable starts FALSE; the home is commanded explicitly in the test flow.
IF bStagesInit THEN
    FOR nInit := 1 TO 5 DO
        afbStage[nInit].SetModeEnableLimits(
            LimBackward    := TRUE,
            LimForward     := TRUE,
            HomeEnable     := FALSE,
            BrakeMode      := E_StageBrakeMode.IF_ENABLED,
            EnableMode     := E_StageEnableMode.ALWAYS,
            HomeMode       := E_EpicsHomeCmd.LOW_LIMIT,
            UserEnable     := TRUE,
            HardwareEnable := TRUE);
    END_FOR
    bStagesInit := FALSE;
END_IF

T01_HomeThenCenterThenZero();
T02_CenterOffset_Y_Geometry();
T03_UserEnableDrop_RedirectsToError();
T04_ReHome_ReArmsFromIdle();
T05_NoHomingEdge_StaysIdle();

// Integration: drive a real limit-switch home (cam-switch pulser pattern, as in
// the T10 reference), with FB_HomeToCenter observing the NC home and performing the
// centering move + MC_SetPosition zero. Asserts the real axis is homed and that
// NcToPlc.ActPos was zeroed at the center position.
METHOD PRIVATE T01_HomeThenCenterThenZero
VAR_INST
    fbUUT : FB_HomeToCenter(iMotionStage := afbStage[1])
            := (fCenterOffset := 2.5, fDefaultVelocity := 10.0);
    fbSearch    : TON := (PT := T#5000MS);
    fbSync      : TON := (PT := T#5000MS);
    fbTimeout   : TON := (IN := TRUE, PT := T#120S);
    nStep       : INT;
END_VAR
// Drive the simulated limit-switch home (mirrors T10); FB observes alongside
CASE nStep OF
0:  // wait for the stage to come ready before commanding anything
    IF afbStage[1].stMotionStatus.bStageReady THEN
        nStep := 1;
    END_IF

1:  // NC-side command of the low-limit home; FB will see bHoming rise
    // afbStage[1].MotionCmd.eHomeMode --> fixed on newer releases, cant be used now
    afbStage[1].Home(HomePosition := 20.0, HomeMode := E_EpicsHomeCmd.LOW_LIMIT);
    fbSearch.IN := TRUE;
    nStep := 2;

2:  // search phase: forward-only to find the switch
    IF fbSearch.Q THEN
        afbStage[1].EnableLimits(BackwardEnable := FALSE, ForwardEnable := TRUE, HomeEnable := FALSE);
        fbSearch.IN := FALSE;
        fbSync.IN   := TRUE;
        nStep := 3;
    END_IF

3:  // sync phase: re-enable both; home completes -> bDone AND bHomed
    IF fbSync.Q THEN
        afbStage[1].EnableLimits(BackwardEnable := TRUE, ForwardEnable := TRUE, HomeEnable := FALSE);
        fbSync.IN := FALSE;
        nStep := 4;
    END_IF

4:  // home complete: the FB should have observed bHoming->(bDone AND bHomed) and be
    //  centering (CenterMove) or already zeroing (WaitCenterDone) or finished.
    IF afbStage[1].stMotionStatus.bDone AND afbStage[1].stMotionStatus.bHomed THEN
        nStep := 5;
    END_IF

5:  // wait for the FB to finish its own center + zero sequence
    IF fbUUT.bCentered AND fbUUT.bHomeDone THEN
        nStep := 6;
    END_IF

6: ;   // terminal - asserts below
END_CASE

//  All sub-FBs ticked unconditionally outside the CASE, stage last so the FB
//  reads current-cycle status.
fbSearch();
fbSync();
fbTimeout();
afbStage[1]();
fbUUT();

//  Terminal / timeout
TEST('T01_HomeThenCenterThenZero');
IF nStep = 6 THEN
    AssertTrue(
        Condition := fbAxisRef[1].Status.Homed,
        Message   := 'T01: axis should be homed');
    AssertTrue(
        Condition := fbUUT.bCentered,
        Message   := 'T01: FB should report centered');
    //  MC_SetPosition zeroed the centered position -> ActPos ~ 0
    AssertEquals_LREAL(
        Expected := 0.0,
        Actual   := fbAxisRef[1].NcToPlc.ActPos,
        Delta    := 0.01,
        Message  := 'T01: position should be zeroed at center by MC_SetPosition');
    TEST_FINISHED();
ELSIF fbTimeout.Q THEN
    AssertTrue(
        Condition := FALSE,
        Message   := CONCAT('T01: timed out at step ', TO_STRING(nStep)));
    TEST_FINISHED();
END_IF
END_METHOD

// Happy path with the Y center offset (6.5) to confirm fCenterOffset is honored
// and the axis is zeroed at center by MC_SetPosition.
METHOD PRIVATE T02_CenterOffset_Y_Geometry
VAR_INST
    fbUUT : FB_HomeToCenter(iMotionStage := afbStage[2])
            := (fCenterOffset := 6.5, fDefaultVelocity := 10.0);
    fbSearch  : TON := (PT := T#5000MS);
    fbSync    : TON := (PT := T#5000MS);
    fbTimeout : TON := (IN := TRUE, PT := T#120S);
    nStep     : INT;
END_VAR
CASE nStep OF
0:  IF afbStage[2].stMotionStatus.bStageReady THEN
        nStep := 1;
    END_IF

1:  afbStage[2].Home(HomePosition := 20.0, HomeMode := E_EpicsHomeCmd.LOW_LIMIT);
    fbSearch.IN := TRUE;
    nStep := 2;

2:  IF fbSearch.Q THEN
        afbStage[2].EnableLimits(BackwardEnable := FALSE, ForwardEnable := TRUE, HomeEnable := FALSE);
        fbSearch.IN := FALSE;
        fbSync.IN   := TRUE;
        nStep := 3;
    END_IF

3:  IF fbSync.Q THEN
        afbStage[2].EnableLimits(BackwardEnable := TRUE, ForwardEnable := TRUE, HomeEnable := FALSE);
        fbSync.IN := FALSE;
        nStep := 4;
    END_IF

4:  IF afbStage[2].stMotionStatus.bDone AND afbStage[2].stMotionStatus.bHomed THEN
        nStep := 5;
    END_IF

5:  IF fbUUT.bCentered AND fbUUT.bHomeDone THEN
        nStep := 6;
    END_IF

6: ;
END_CASE

fbSearch();
fbSync();
fbTimeout();
afbStage[2]();
fbUUT();

TEST('T02_CenterOffset_Y_Geometry');
IF nStep = 6 THEN
    AssertTrue(
        Condition := fbAxisRef[2].Status.Homed,
        Message   := 'T02: axis should be homed');
    AssertEquals_LREAL(
        Expected := 0.0,
        Actual   := fbAxisRef[2].NcToPlc.ActPos,
        Delta    := 0.01,
        Message  := 'T02: position should be zeroed at center (offset 6.5) by MC_SetPosition');
    TEST_FINISHED();
ELSIF fbTimeout.Q THEN
    AssertTrue(Condition := FALSE,
        Message := CONCAT('T02: timed out at step ', TO_STRING(nStep)));
    TEST_FINISHED();
END_IF
END_METHOD

// Dropping UserEnable mid-home faults the stage (bError, bStageReady still TRUE
// as a boot flag) -> FB redirects to Error, latches bLocalError, never centers.
METHOD PRIVATE T03_UserEnableDrop_RedirectsToError
VAR_INST
    fbUUT : FB_HomeToCenter(iMotionStage := afbStage[3])
            := (fCenterOffset := 2.5, fDefaultVelocity := 10.0);
    fbSearch  : TON := (PT := T#5000MS);
    fbSync    : TON := (PT := T#5000MS);
    fbTimeout : TON := (IN := TRUE, PT := T#120S);
    nStep     : INT;
END_VAR
CASE nStep OF
0:  IF afbStage[3].stMotionStatus.bStageReady THEN
        nStep := 1;
    END_IF

1:  // command the home so the FB enters its sequence
    afbStage[3].Home(HomePosition := 20.0, HomeMode := E_EpicsHomeCmd.LOW_LIMIT);
    fbSearch.IN := TRUE;
    nStep := 2;

2:  // mid-home, pull user-enable: faults the stage. bStageReady is a boot flag and
    //  stays TRUE, so rtError (bError AND bStageReady) fires in the FB.
    IF fbSearch.Q THEN
        afbStage[3].SetModeEnableLimits(
            LimBackward    := TRUE,
            LimForward     := TRUE,
            HomeEnable     := FALSE,
            BrakeMode      := E_StageBrakeMode.IF_ENABLED,
            EnableMode     := E_StageEnableMode.ALWAYS,
            HomeMode       := E_EpicsHomeCmd.LOW_LIMIT,
            UserEnable     := FALSE,
            HardwareEnable := TRUE);
        nStep := 3;
    END_IF

3:  // wait for the FB to redirect to Error
    IF fbUUT.eHomeCenterState = E_HomeCenterState.Error THEN
        nStep := 6;
    END_IF
END_CASE

fbSearch();
fbSync();
fbTimeout();
afbStage[3]();
fbUUT();

TEST('T03_UserEnableDrop_RedirectsToError');
IF nStep = 6 THEN
    AssertEquals_INT(
        Expected := E_HomeCenterState.Error,
        Actual   := fbUUT.eHomeCenterState,
        Message  := 'T03: dropping UserEnable should redirect FB to Error');
    AssertTrue(
        Condition := fbUUT.bLocalError,
        Message   := 'T03: bLocalError should latch in Error');
    AssertFalse(
        Condition := fbUUT.bCentered,
        Message   := 'T03: must NOT report centered after an error');
    AssertFalse(
        Condition := fbUUT.bHomeDone,
        Message   := 'T03: must NOT report home done after an error');
    TEST_FINISHED();
ELSIF fbTimeout.Q THEN
    AssertTrue(Condition := FALSE,
        Message := CONCAT('T03: timed out at step ', TO_STRING(nStep)));
    TEST_FINISHED();
END_IF
END_METHOD

// Complete one home+center cycle, confirm the FB returns to Idle, then command a
// second home and confirm it re-arms and re-zeroes (HomingDone -> Idle re-arm path).
METHOD PRIVATE T04_ReHome_ReArmsFromIdle
VAR_INST
    fbUUT : FB_HomeToCenter(iMotionStage := afbStage[4])
            := (fCenterOffset := 2.5, fDefaultVelocity := 10.0);
    fbSearch  : TON := (PT := T#5000MS);
    fbSync    : TON := (PT := T#5000MS);
    fbTimeout : TON := (IN := TRUE, PT := T#120S);
    nStep     : INT;
    bFirstDone : BOOL;
END_VAR
CASE nStep OF
0:  IF afbStage[4].stMotionStatus.bStageReady THEN
        nStep := 1;
    END_IF

1:  afbStage[4].Home(HomePosition := 20.0, HomeMode := E_EpicsHomeCmd.LOW_LIMIT);
    fbSearch.IN := TRUE;
    nStep := 2;

2:  IF fbSearch.Q THEN
        afbStage[4].EnableLimits(BackwardEnable := FALSE, ForwardEnable := TRUE, HomeEnable := FALSE);
        fbSearch.IN := FALSE;
        fbSync.IN   := TRUE;
        nStep := 3;
    END_IF

3:  IF fbSync.Q THEN
        afbStage[4].EnableLimits(BackwardEnable := TRUE, ForwardEnable := TRUE, HomeEnable := FALSE);
        fbSync.IN := FALSE;
        nStep := 4;
    END_IF

4:  IF afbStage[4].stMotionStatus.bDone AND afbStage[4].stMotionStatus.bHomed THEN
        nStep := 5;
    END_IF

5:  // first cycle complete; confirm FB returned to Idle (re-armable)
    IF fbUUT.bCentered AND fbUUT.bHomeDone THEN
        bFirstDone := TRUE;
        nStep := 6;
    END_IF

6:  // FB should restore params and fall back to Idle on its own
    IF fbUUT.eHomeCenterState = E_HomeCenterState.Idle THEN
        nStep := 7;
    END_IF

7:  // re-home: command Home() again, re-run the pulser dance
    afbStage[4].Home(HomePosition := 20.0, HomeMode := E_EpicsHomeCmd.LOW_LIMIT);
    fbSearch.IN := TRUE;
    nStep := 8;

8:  IF fbSearch.Q THEN
        afbStage[4].EnableLimits(BackwardEnable := FALSE, ForwardEnable := TRUE, HomeEnable := FALSE);
        fbSearch.IN := FALSE;
        fbSync.IN   := TRUE;
        nStep := 9;
    END_IF

9:  IF fbSync.Q THEN
        afbStage[4].EnableLimits(BackwardEnable := TRUE, ForwardEnable := TRUE, HomeEnable := FALSE);
        fbSync.IN := FALSE;
        nStep := 10;
    END_IF

10: IF fbUUT.bCentered AND fbUUT.bHomeDone THEN
        nStep := 11;
    END_IF

11: ;
END_CASE

fbSearch();
fbSync();
fbTimeout();
afbStage[4]();
fbUUT();

TEST('T04_ReHome_ReArmsFromIdle');
IF nStep = 11 THEN
    AssertTrue(
        Condition := bFirstDone,
        Message   := 'T04: first home/center cycle should have completed');
    AssertTrue(
        Condition := fbUUT.bCentered,
        Message   := 'T04: second home/center cycle should re-arm and complete');
    AssertEquals_LREAL(
        Expected := 0.0,
        Actual   := fbAxisRef[4].NcToPlc.ActPos,
        Delta    := 0.01,
        Message  := 'T04: position should be re-zeroed after the second cycle');
    TEST_FINISHED();
ELSIF fbTimeout.Q THEN
    AssertTrue(Condition := FALSE,
        Message := CONCAT('T04: timed out at step ', TO_STRING(nStep)));
    TEST_FINISHED();
END_IF
END_METHOD

// With no home commanded, bHoming never rises -> FB must remain Idle and never
// center (rising-edge entry, not level)
METHOD PRIVATE T05_NoHomingEdge_StaysIdle
VAR_INST
    fbUUT : FB_HomeToCenter(iMotionStage := afbStage[5])
            := (fCenterOffset := 2.5, fDefaultVelocity := 10.0);
    fbSettle  : TON := (PT := T#2000MS);
    fbTimeout : TON := (IN := TRUE, PT := T#30S);
    nStep     : INT;
END_VAR
CASE nStep OF
0:  IF afbStage[5].stMotionStatus.bStageReady THEN
        nStep := 1;
    END_IF

1:  // never command a home -> bHoming never rises. Let the stage idle for a while.
    fbSettle.IN := TRUE;
    nStep := 2;

2:  IF fbSettle.Q THEN
        nStep := 6;
    END_IF
END_CASE

fbSettle();
fbTimeout();
afbStage[5]();
fbUUT();

TEST('T05_NoHomingEdge_StaysIdle');
IF nStep = 6 THEN
    AssertEquals_INT(
        Expected := E_HomeCenterState.Idle,
        Actual   := fbUUT.eHomeCenterState,
        Message  := 'T05: with no bHoming edge the FB must stay Idle');
    AssertFalse(
        Condition := fbUUT.bCentered,
        Message   := 'T05: must not center without a home');
    TEST_FINISHED();
ELSIF fbTimeout.Q THEN
    AssertTrue(Condition := FALSE,
        Message := CONCAT('T05: timed out at step ', TO_STRING(nStep)));
    TEST_FINISHED();
END_IF
END_METHOD

END_FUNCTION_BLOCK

// ---- POUs/FB_HomeToCenter.TcPOU
(*  FB_HomeToCenter - Limit-switch homing + centering sequence.

 Overview:
   This FB does NOT command the home; it observes the rising edge of bHoming, waits for the
   drive to confirm bDone AND bHomed, then issues a centering AbsoluteMove to
   fCenterOffset and zeroes the position via MC_SetPosition.the drive's own switch-homing finds the reference, so the FB only sequences
   "wait homed -> center -> zero".

 Per-instance wiring (via FB_Init):
   iMotionStage : the stage interface this FB sequences.
   refAxis      : the AXIS_REF used for the position-zero (e.g. GVL_AXES.Axes[2]
                  for X, GVL_AXES.Axes[3] for Y).

 Per-instance parameters:
   fCenterOffset    : centering target after home (X: 2.5, Y: 6.5).
   fDefaultVelocity : centering move velocity, also the velocity restore fallback.
*)
FUNCTION_BLOCK FB_HomeToCenter
VAR_INPUT
    fCenterOffset    : LREAL;
    fDefaultVelocity : LREAL;
END_VAR
VAR
    iMotionStage : I_MotionStage;

    {attribute 'hide'}
    rtHomingStart  : R_TRIG;
    {attribute 'hide'}
    rtWaitHomeDone : R_TRIG;
    {attribute 'hide'}
    rtCenterDone   : R_TRIG;
    {attribute 'hide'}
    rtError        : R_TRIG;

    fPrevVelocity   : LREAL;
    fbMcSetPosition : MC_SetPosition;
END_VAR
VAR_OUTPUT
    {attribute 'pytmc' := '
        pv: bCentered
        io: i
        field: ZNAM FALSE
        field: ONAM TRUE
        field: DESC TRUE if the stage is centered
    '}
    bCentered      : BOOL;
    bHomeDone      : BOOL;
    bLocalError    : BOOL;
    eHomeCenterState : E_HomeCenterState := E_HomeCenterState.Idle;
END_VAR

IF (iMotionStage = 0) THEN
    RETURN;
END_IF

// Edge detection - all R_TRIG instances tick every cycle, outside the CASE.
rtError(CLK := iMotionStage.MotionStatus.bError AND iMotionStage.MotionStatus.bStageReady);
rtHomingStart(CLK := iMotionStage.MotionStatus.bHoming);
// Fires when the drive confirms both done and homed during the wait state.
rtWaitHomeDone(CLK := iMotionStage.MotionStatus.bDone
        AND iMotionStage.MotionStatus.bHomed
        AND (eHomeCenterState = E_HomeCenterState.WaitHomeDone));
// Fires when the centering move completes.
rtCenterDone(CLK := iMotionStage.MotionStatus.bDone
        AND (eHomeCenterState = E_HomeCenterState.CenterMove));

// Any drive error redirects to Error from any point in the sequence.
IF rtError.Q THEN
    eHomeCenterState := E_HomeCenterState.Error;
END_IF

CASE eHomeCenterState OF
    E_HomeCenterState.Idle:
        // The NC side owns the home trigger. Enter the sequence on the rising
        // edge of bHoming (NC is the source of truth).
        IF rtHomingStart.Q THEN
            Reset();
            bCentered := FALSE;
            // Preserve current velocity to restore after centering; fall back to default.
            IF iMotionStage.MotionCmd.fVelocity <> 0.0 THEN
                fPrevVelocity := iMotionStage.MotionCmd.fVelocity;
            ELSE
                fPrevVelocity := fDefaultVelocity;
            END_IF
            eHomeCenterState := E_HomeCenterState.WaitHomeDone;
        END_IF

    E_HomeCenterState.WaitHomeDone:
        // Drive is homing against the switch. Wait for both bDone and bHomed,
        // confirming the homing move has fully settled, then center.
        IF rtWaitHomeDone.Q THEN
            iMotionStage.AbsoluteMoveDefault(
                Position := fCenterOffset,
                Velocity := fDefaultVelocity
            );
            eHomeCenterState := E_HomeCenterState.CenterMove;
        END_IF

    E_HomeCenterState.CenterMove:
        // AbsoluteMoveDefault clears bDone before starting, so rtCenterDone only
        // fires on the fresh rising edge from THIS move completing.
        IF rtCenterDone.Q THEN
            // Define the current (centered) position as zero.
            fbMcSetPosition.Execute := TRUE;
            eHomeCenterState := E_HomeCenterState.WaitCenterDone;
        END_IF

    E_HomeCenterState.WaitCenterDone:
        // fbMcSetPosition runs unconditionally below the CASE each cycle.
        IF fbMcSetPosition.Done THEN
            fbMcSetPosition.Execute := FALSE;
            bCentered := TRUE;
            bHomeDone := TRUE;
            eHomeCenterState := E_HomeCenterState.HomingDone;
        END_IF

    E_HomeCenterState.HomingDone:
        // Restore motion parameters to the pre-homing state, then return to Idle
        // ready for the next NC-initiated homing cycle.
        iMotionStage.SetDefaultMotionParameters(
            HomePosition := 0.0,
            Velocity     := fPrevVelocity
        );
        iMotionStage.MotionCmd.fPosition := iMotionStage.MotionCmd.fHomePosition;
        eHomeCenterState := E_HomeCenterState.Idle;

    E_HomeCenterState.Error:
        // Latch error output and safe the sequence. Caller must invoke Reset().
        bLocalError := TRUE;
        fbMcSetPosition.Execute := FALSE;
        bCentered := FALSE;
        bHomeDone := FALSE;
        IF iMotionStage.ExMotionStatus.bLatchReset THEN
            bLocalError := FALSE;
            eHomeCenterState := E_HomeCenterState.Idle;
        END_IF

END_CASE

// MC_SetPosition runs every cycle; Execute is gated by WaitCenterDone above.
// Axis comes from the injected refAxis so X and Y target their own axes.
fbMcSetPosition(
    Axis     := iMotionStage.Axis,
    Mode     := 0,
    Position := 0.0
);

//FB_Init is always available implicitly and it is used primarily for initialization.
//The return value is not evaluated. For a specific influence, you can also declare the
//methods explicitly and provide additional code there with the standard initialization
//code. You can evaluate the return value.
METHOD FB_Init: BOOL
VAR_INPUT
    bInitRetains: BOOL; // TRUE: the retain variables are initialized (reset warm / reset cold)
    bInCopyCode: BOOL;  // TRUE: the instance will be copied to the copy code afterward (online change)
    iMotionStage : I_MotionStage;
END_VAR
THIS^.iMotionStage := iMotionStage;
END_METHOD

METHOD Reset
VAR_INPUT
END_VAR
bCentered := FALSE;
bHomeDone := FALSE;
bLocalError := FALSE;
fbMcSetPosition.Execute := FALSE;
eHomeCenterState := E_HomeCenterState.Idle;
END_METHOD

END_FUNCTION_BLOCK

// ---- POUs/PRG_XY.TcPOU
PROGRAM PRG_XY
VAR
     {attribute 'pytmc' := '
        axis-link: GVL_Axes.Axes[2]
        pv: SH1L2:PP:MMS:02
    '}
    {attribute 'TcLinkTo' := '.fbLimSwStatus.bLimitFwd  := TIIB[XY]^DI Inputs Channel 1^Input 2;
                              .fbLimSwStatus.bLimitBwd := TIIB[XY]^DI Inputs Channel 1^Input 1;
                              .fbEncoderScaling.nRawEncoderUDINT  := TIIB[XY]^FB Position Channel 1^Position'}
    fbX : FB_MotionStageNC(
        sName                  := 'PP_X',
        AxisRef                := GVL_Axes.Axes[2],
        iPersistentDataStorage := GVL_Common.fbPersistentDataStorage
    ) := (HomeMode := E_EpicsHomeCmd.LOW_LIMIT);

    {attribute 'pytmc' := '
        axis-link: GVL_Axes.Axes[3]
        pv: SH1L2:PP:MMS:03
    '}
    {attribute 'TcLinkTo' := '.fbLimSwStatus.bLimitFwd  := TIIB[XY]^DI Inputs Channel 2^Input 1;
                              .fbLimSwStatus.bLimitBwd := TIIB[XY]^DI Inputs Channel 2^Input 2;
                              .fbEncoderScaling.nRawEncoderUDINT  := TIIB[XY]^FB Position Channel 2^Position'}
    fbY : FB_MotionStageNC(
        sName                  := 'PP_Y',
        AxisRef                := GVL_Axes.Axes[3],
        iPersistentDataStorage := GVL_Common.fbPersistentDataStorage
    ) := (HomeMode := E_EpicsHomeCmd.LOW_LIMIT);

    {attribute 'pytmc' := '
        pv: SH1L2:PP:MMS:02
    '}
    fbXEPS : LCLS_MotionAbstraction.FB_EPS;

    {attribute 'pytmc' := '
        pv: SH1L2:PP:MMS:03
    '}
    fbYEPS : LCLS_MotionAbstraction.FB_EPS;

    {attribute 'pytmc' := '
        pv: SH1L2:PP:MMS
    '}
    fbPPEPS : FB_PPEPS (
        iXEPS  := fbXEPS,
        iYEPS  := fbYEPS,
        iXMotionStage:=fbX,
        iYMotionStage:=fbY
    );
    {attribute 'pytmc' := '
        pv: SH1L2:PP:MMS:02
    '}
    fbXHome : FB_HomeToCenter(
        iMotionStage:=fbX
    );
    {attribute 'pytmc' := '
        pv: SH1L2:PP:MMS:03
    '}
    fbYHome : FB_HomeToCenter(iMotionStage:=fbY);
    bInit   : BOOL := TRUE;

END_VAR

VAR PERSISTENT
    {attribute 'pytmc' := '
        pv: SH1L2:PP:MMS:02:fXCenterOffset
        io: io
        field: DESC Centering Offset
    '}
    fXCenterOffset: LREAL := 2.5;

    {attribute 'pytmc' := '
        pv: SH1L2:PP:MMS:03:fYCenterOffset
        io: io
        field: DESC Centering Offset
    '}
    fYCenterOffset: LREAL := 6.5;

    {attribute 'pytmc' := '
        pv: SH1L2:PP:MMS:03:fInOutThrsh
        io: io
        field: DESC In/Out Threshold
    '}
    fInOutThrsh : LREAL;

    {attribute 'pytmc' := '
        pv: SH1L2:PP:MMS:03:eInOutStatus
        io: i
        field: DESC In/Out Status
    '}
    eInOutStatus : E_PPStatus;
END_VAR

IF bInit THEN
    fbX.AssignEPS(iEPS:=fbXEPS);
    fbX.SetModeEnableLimits(
        LimBackward     := TRUE,
        LimForward      := TRUE,
        HomeEnable      := FALSE,
        BrakeMode       := E_StageBrakeMode.IF_ENABLED,
        EnableMode      := E_StageEnableMode.DURING_MOTION,
        HomeMode        := 1,
        UserEnable      := TRUE,
        HardwareEnable  := TRUE
    );
    fbX.SetDefaultMotionParameters (
        HomePosition    := 0.0,
        Velocity        := 3.0,
    );
    // Y
    fbY.AssignEPS(iEPS:=fbYEPS);
    fbY.SetModeEnableLimits(
        LimBackward     := TRUE,
        LimForward      := TRUE,
        HomeEnable      := FALSE,
        BrakeMode       := E_StageBrakeMode.IF_ENABLED,
        EnableMode      := E_StageEnableMode.DURING_MOTION,
        HomeMode        := 1,
        UserEnable      := TRUE,
        HardwareEnable  := TRUE
    );
    fbY.SetDefaultMotionParameters (
        HomePosition    := 0.0,
        Velocity        := 4.0,
    );
   bInit := FALSE;
END_IF

fbPPEPS(
    bPickActive := GVL_Common.eModeSelect <> E_ModeSelector.ModeNone
);

fbX();
fbXHome(
    fCenterOffset    := fXCenterOffset,
    fDefaultVelocity := fbX.MotionCmd.fVelocity
);

fbY();
fbYHome(
    fCenterOffset    := fYCenterOffset,
    fDefaultVelocity := fbY.MotionCmd.fVelocity
);

// Pulse Picker status (Given Y axis moving up is from 0-20.1mm)
IF NOT fbY.MotionStatus.bMoving THEN
    IF fbY.MotionStatus.fActPosition > fInOutThrsh THEN
        eInOutStatus := E_PPStatus.OUT;
    ELSE
        eInOutStatus := E_PPStatus.IN;
    END_IF
ELSE
    eInOutStatus := E_PPStatus.UNKNOWN;
END_IF

END_PROGRAM

// ---- POUs/PRG_S.TcPOU
PROGRAM PRG_S
VAR
    {attribute 'pytmc' := '
        pv: SH1L2:PP:MMS:01:eModeSelector
        io: io
        field: DESC Pulse Picker mode selector
    '}
    eModeReq    : E_ModeSelector := E_ModeSelector.ModeNone;
    eStatus     : E_StatusIndicator;
    ePickState  : E_PickerState := E_PickerState.Init;
    eState      : INT := 0;

    {attribute 'pytmc' := '
        axis-link: GVL_Axes.Axes[1]
        pv: SH1L2:PP:MMS:01
    '}
    {attribute 'TcLinkTo' := '.fbEncoderScaling.nRawEncoderUDINT := TIIB[Spindle]^FB Position Channel 1^Position'}
    fbS : FB_MotionStageNC(
        sName    := 'Spindle',
        AxisRef  := GVL_Axes.Axes[1],
        iPersistentDataStorage := GVL_Common.fbPersistentDataStorage
    ) := (HomeMode := E_EpicsHomeCmd.HOME_INDEX);

    {attribute 'pytmc' := '
        pv: SH1L2:PP:MMS:01
    '}
    fbTrigMgr : FB_TriggerSetpointManager(
        AxisRef      := GVL_Axes.Axes[1],
        iMotionStage := fbS
    );

    nErrCode : INT := 0;

    fbMoveNearest : FB_MoveToNearestClosed(iMotionStage := fbS);
    fbFastOpen    : FB_FastOpen(iMotionStage := fbS);
    fbFastClose   : FB_FastClose(iMotionStage := fbS);

    {attribute 'pytmc' := '
        pv: SH1L2:PP:MMS:01
    '}
    fbHomeIdx : FB_SpindleHomeToCenter(iMotionStage := fbS);

    bPicking   : BOOL;
    ftStopPick : F_TRIG;

END_VAR

VAR PERSISTENT
    {attribute 'pytmc' := '
        pv: SH1L2:PP:MMS:01:fCenterOffset
        io: io
        field: DESC Center Position Offset
    '}
    fCenterOffset : LREAL := 113.247;

    {attribute 'pytmc' := '
        pv: SH1L2:PP:MMS:01:fStopPos
        io: io
        field: DESC End Stop Positive
    '}
    fStopPos : LREAL := 11.25;

    {attribute 'pytmc' := '
        pv: SH1L2:PP:MMS:01:fStopNeg
        io: io
        field: DESC End Stop Negative
    '}
    fStopNeg : LREAL := -12.5;

    {attribute 'pytmc' := '
        pv: SH1L2:PP:MMS:01:fCenter
        io: io
        field: DESC Center Position
    '}
    fCenter : LREAL := 0.0;

    fDefVel : LREAL := 1650;
END_VAR

CASE ePickState OF

    // INIT ALL
    E_PickerState.Init:
        fbS.SetModeEnableLimits(
            LimBackward    := TRUE,
            LimForward     := TRUE,
            HomeEnable     := FALSE,
            BrakeMode      := E_StageBrakeMode.IF_ENABLED,
            EnableMode     := E_StageEnableMode.ALWAYS,
            HomeMode       := E_EpicsHomeCmd.HOME_INDEX,
            UserEnable     := TRUE,
            HardwareEnable := TRUE
        );
        fbS.SetDefaultMotionParameters(
            HomePosition := 0.0,
            Velocity     := fDefVel,
        );

        // Enable backlash (negative) compensation
        fbS.BacklashCompensation(Enable:=TRUE, RampVelo:=fDefVel/10.0);
        // the backlash value provided here is from demo (must be adapted for prod)
        fbTrigMgr.Reset();
        GVL_Common.eModeSelect := E_ModeSelector.ModeNone;
        ePickState := E_PickerState.ModeSelect;

    // WAIT USER MODE SELECT
    E_PickerState.ModeSelect:
        bPicking := FALSE;
        fbTrigMgr.Stop();
        IF fbS.MotionStatus.bError THEN
            ePickState := E_PickerState.ErrorState;
        ELSIF eModeReq <> E_ModeSelector.ModeNone THEN
            GVL_Common.eModeSelect := eModeReq;
            eStatus    := E_StatusIndicator.Init;
            ePickState := E_PickerState.ModeExecute;
        END_IF

    // MAIN MODE EXECUTE
    E_PickerState.ModeExecute:
        CASE GVL_Common.eModeSelect OF
            E_ModeSelector.FlipFlop, E_ModeSelector.Burst:
                CASE eStatus OF
                    E_StatusIndicator.Init:
                        bPicking := TRUE;
                        fbTrigMgr.Stop();
                        IF fbS.MotionStatus.bPowerIsEnabled THEN
                            fbMoveNearest.Start();
                        END_IF
                        eStatus := E_StatusIndicator.Closed;

                    E_StatusIndicator.Closed:
                        IF fbMoveNearest.Closed THEN
                            fbTrigMgr.Start();
                            eStatus := E_StatusIndicator.Wait;
                        END_IF

                    E_StatusIndicator.Wait:
                        IF eModeReq = E_ModeSelector.ModeNone THEN
                            eStatus    := E_StatusIndicator.Init;
                            GVL_Common.eModeSelect := E_ModeSelector.ModeNone;
                            ePickState := E_PickerState.ModeSelect;
                        ELSIF eModeReq = E_ModeSelector.Close THEN
                            fbTrigMgr.Stop();
                            GVL_Common.eModeSelect := E_ModeSelector.Close;
                            eStatus    := E_StatusIndicator.Init;
                            ePickState := E_PickerState.ModeExecute;
                        ELSIF eModeReq = E_ModeSelector.Open THEN
                            fbTrigMgr.Stop();
                            GVL_Common.eModeSelect := E_ModeSelector.Open;
                            eStatus    := E_StatusIndicator.Init;
                            ePickState := E_PickerState.ModeExecute;
                        END_IF
                END_CASE

            E_ModeSelector.Close:
                CASE eStatus OF
                    E_StatusIndicator.Init:
                        fbFastClose.Start();
                        eStatus := E_StatusIndicator.Closed;
                    E_StatusIndicator.Closed:
                        IF fbFastClose.Closed THEN
                            eModeReq	:= E_ModeSelector.ModeNone;
                            GVL_Common.eModeSelect := E_ModeSelector.ModeNone;
                            eStatus    := E_StatusIndicator.Init;
                            ePickState := E_PickerState.ModeSelect;
                        END_IF
                END_CASE

            E_ModeSelector.Open:
                CASE eStatus OF
                    E_StatusIndicator.Init:
                        fbFastOpen.Start();
                        eStatus := E_StatusIndicator.Opened;
                    E_StatusIndicator.Opened:
                        IF fbFastOpen.Opened THEN
                            eModeReq	:= E_ModeSelector.ModeNone;
                            GVL_Common.eModeSelect := E_ModeSelector.ModeNone;
                            eStatus    := E_StatusIndicator.Init;
                            ePickState := E_PickerState.ModeSelect;
                        END_IF
                END_CASE

            E_ModeSelector.Home:
                CASE eStatus OF
                    E_StatusIndicator.Init:
                        IF fbS.MotionStatus.bMoving THEN
                            fbS.Halt();
                        END_IF
                        eStatus := E_StatusIndicator.Closed;
                    E_StatusIndicator.Closed:
                        IF fbS.MotionStatus.bDone OR NOT fbS.MotionStatus.bMoving THEN
                            fbS.Home(
                                HomePosition := 0.0,
                                HomeMode     := E_EPicsHomeCmd.HOME_INDEX
                            );
                            eStatus := E_StatusIndicator.Done;
                        END_IF
                    E_StatusIndicator.Done:
                        IF fbHomeIdx.bCentered THEN
                            eModeReq               := E_ModeSelector.ModeNone;
                            GVL_Common.eModeSelect := E_ModeSelector.ModeNone;
                            eStatus    := E_StatusIndicator.Init;
                            ePickState := E_PickerState.ModeSelect;
                        END_IF
                END_CASE

            ELSE
                eStatus                := E_StatusIndicator.Init;
                GVL_Common.eModeSelect := E_ModeSelector.ModeNone;
                ePickState             := E_PickerState.ModeSelect;
        END_CASE

    E_PickerState.ErrorState:
        fbTrigMgr.Stop();
        IF NOT fbS.MotionStatus.bError THEN
            ePickState := E_PickerState.ModeSelect;
        END_IF

    ELSE
        ePickState := E_PickerState.Init;
END_CASE

// Global reset / halt overrides
IF fbS.MotionCmd.bReset THEN
    fbTrigMgr.Reset();
    fbHomeIdx.Reset();
    fbS.ExMotionStatus.bLatchReset := FALSE;
    eModeReq               := E_ModeSelector.ModeNone;
    GVL_Common.eModeSelect := E_ModeSelector.ModeNone;
    eStatus    := E_StatusIndicator.Init;
    ePickState := E_PickerState.ModeSelect;
ELSIF fbS.MotionCmd.bHalt AND (GVL_Common.eModeSelect <> E_ModeSelector.Home) THEN
    fbTrigMgr.Stop();
    eModeReq               := E_ModeSelector.ModeNone;
    GVL_Common.eModeSelect := E_ModeSelector.ModeNone;
    eStatus    := E_StatusIndicator.Init;
    ePickState := E_PickerState.ModeSelect;
END_IF

fbTrigMgr(
    Mode := eModeReq,
    fStopPos:=fStopPos,
    fStopNeg:=fStopNeg,
    fCenter:=fCenter
);

fbMoveNearest();

fbFastOpen(
    fCenter:=fCenter
);

fbFastClose(
    fStopPos:=fStopPos
);

fbHomeIdx(
    fCenterOffset    := fCenterOffset,
    fDefaultVelocity := fDefVel
);

fbS();
IF fbS.MotionStatus.bError AND fbS.MotionStatus.bStageReady THEN
    ePickState := E_PickerState.ErrorState;
END_IF

END_PROGRAM

// ---- POUs/FB_TriggerSetpointManager.TcPOU
FUNCTION_BLOCK FB_TriggerSetpointManager
VAR_INPUT
    Mode     : E_ModeSelector;
    bWaitDone : BOOL := TRUE;
    fStopPos : LREAL;
    fStopNeg : LREAL;
    fCenter : LREAL;
END_VAR

VAR_OUTPUT
    fSetpoint : LREAL;
    nMoveIdx  : INT;
    bBusy     : BOOL;
END_VAR

VAR
    fbMoveAbs0 : MC_MoveAbsolute;
    fbMoveAbs1 : MC_MoveAbsolute;
    AxisRef    : REFERENCE TO AXIS_REF;
    iMotionStage : I_MotionStage;

    fbTrigSrc  : LCLS_Tc_MotSync.FB_TriggerSourceEL1124;
    {attribute 'pytmc' := 'pv:'}
    fbTrigMgr  : LCLS_Tc_MotSync.FB_TriggerManagerEL1124(
        fTriggerFrequencyExpected := fTargetFreq,
        iTriggerSource := fbTrigSrc
    );

    eState       : INT := 0;
    lastEndPoint : LREAL := 0.0;
    bStarted     : BOOL;

    // Overshoot counters
    {attribute 'pytmc' := '
        pv: nOvrCntPos
        io: i
        field: DESC Positive Stop Position over counters
    '}
    nOvrCntPos : UDINT;
    {attribute 'pytmc' := '
        pv: nOvrCntNeg
        io: i
        field: DESC Negative Stop Position over counters
    '}
    nOvrCntNeg : UDINT;

    // Averaging
    bAvg    : BOOL := FALSE;
    fSumPos : LREAL := 0.0;
    nSmpl   : UDINT := 0;
    fAvgPos : LREAL := 0.0;

    rtStop      : R_TRIG;
    rtNewTrig   : R_TRIG;

    // Internal busy flags per FB
    bBusy0 : BOOL;
    bBusy1 : BOOL;

    fTargetFreq : LREAL := 30.0;
    {attribute 'pytmc' := '
        pv: bResetCnt
        io: io
        field: DESC Reset Stop Position over counters
    '}
    bResetCnt  : BOOL := FALSE;
    rtResetCnt : R_TRIG;

END_VAR

VAR PERSISTENT
    {attribute 'pytmc' := '
        pv: fLimitPos
        io: io
        field: DESC Positive Overshoot Limit
    '}
    fLimitPos : LREAL := 14.5;

    {attribute 'pytmc' := '
        pv: fLimitNeg
        io: io
        field: DESC Negative Overshoot Limit
    '}
    fLimitNeg : LREAL := -14.5;
END_VAR

IF iMotionStage = 0 THEN
    RETURN;
END_IF

fbTrigMgr();

// Combine busy flags
bBusy := bBusy0 OR bBusy1;

CASE eState OF
    // WAIT FOR START
    0:
        IF bStarted THEN
            eState := 1;
        END_IF

    // WAIT FOR TRIGGER
    1:
        IF fbTrigMgr.NewTriggerIsAvailable THEN
            // Safety clear of accumulators before a new move
            bAvg    R= FALSE;
            fSumPos := 0.0;
            nSmpl   := 0;
            fAvgPos := 0.0;
            eState  := 2;
        END_IF

    // COMMAND MOVE ON TRIGGER
    2:
        CASE Mode OF
            E_ModeSelector.Burst:
                IF (fSetpoint = fStopPos) OR (fSetpoint = fStopNeg) THEN
                    fSetpoint := fCenter;
                ELSE
                    IF ABS(iMotionStage.MotionStatus.fActPosition - fStopPos)
                      < ABS(iMotionStage.MotionStatus.fActPosition - fStopNeg) THEN
                        fSetpoint := fStopPos;
                    ELSE
                        fSetpoint := fStopNeg;
                    END_IF
                END_IF

            E_ModeSelector.FlipFlop:
                IF lastEndPoint = fStopPos THEN
                    fSetpoint    := fStopNeg;
                    lastEndPoint := fStopNeg;
                ELSE
                    fSetpoint    := fStopPos;
                    lastEndPoint := fStopPos;
                END_IF
        END_CASE

        IF nMoveIdx = 0 THEN
            fbMoveAbs0.Execute := FALSE;
            fbMoveAbs1.Execute := TRUE;
            nMoveIdx := 1;
        ELSE
            fbMoveAbs1.Execute := FALSE;
            fbMoveAbs0.Execute := TRUE;
            nMoveIdx := 0;
        END_IF

        fbTrigMgr.UnlatchTrigger();
        eState := SEL(bWaitDone, 1, 3);

    // WAIT FOR MOVE COMPLETE (optional)
    3:
        IF (nMoveIdx = 0 AND (fbMoveAbs0.Done OR AxisRef.Status.StandStill OR fbMoveAbs0.Error)) OR
           (nMoveIdx = 1 AND (fbMoveAbs1.Done OR AxisRef.Status.StandStill OR fbMoveAbs1.Error)) THEN
            fbMoveAbs0.Execute := FALSE;
            fbMoveAbs1.Execute := FALSE;
            eState := 1;
        END_IF

    ELSE
        eState := 0;
END_CASE

// Motion FBs
fbMoveAbs0(
    Axis       := AxisRef,
    Position   := fSetpoint,
    Velocity   := iMotionStage.MotionCmd.fVelocity,
    BufferMode := MC_BufferMode.MC_Aborting,
    Busy       => bBusy0
);
fbMoveAbs1(
    Axis       := AxisRef,
    Position   := fSetpoint,
    Velocity   := iMotionStage.MotionCmd.fVelocity,
    BufferMode := MC_BufferMode.MC_Aborting,
    Busy       => bBusy1
);

// Detect when stage crosses the setpoint heading toward the stop
rtStop(CLK :=
    (nMoveIdx = 0 AND iMotionStage.MotionStatus.fActPosition < fSetpoint) OR
    (nMoveIdx = 1 AND iMotionStage.MotionStatus.fActPosition > fSetpoint)
);
bAvg S= rtStop.Q;

// Accumulate position while averaging window is open
IF bAvg THEN
    fSumPos := fSumPos + iMotionStage.MotionStatus.fActPosition;
    nSmpl   := nSmpl + 1;
END_IF

// Compute average on the rising edge of the next trigger
// Compute average on the rising edge of the next trigger
rtNewTrig(CLK := fbTrigMgr.NewTriggerIsAvailable);
IF bAvg AND rtNewTrig.Q THEN
    IF nSmpl > 0 THEN
        fAvgPos := fSumPos / nSmpl;
    ELSE
        fAvgPos := iMotionStage.MotionStatus.fActPosition;
    END_IF

    IF fAvgPos > fLimitPos THEN
        nOvrCntPos := nOvrCntPos + 1;
    END_IF
    IF fAvgPos < fLimitNeg THEN
        nOvrCntNeg := nOvrCntNeg + 1;
    END_IF

    fSumPos := 0.0;
    nSmpl   := 0;
    bAvg    := FALSE;
END_IF

// Reset overshoot counters on rising edge, then self-clear
rtResetCnt(CLK := bResetCnt);
IF rtResetCnt.Q THEN
    nOvrCntPos := 0;
    nOvrCntNeg := 0;
    bResetCnt  := FALSE;
END_IF

//FB_Init is always available implicitly and it is used primarily for initialization.
//The return value is not evaluated. For a specific influence, you can also declare the
//methods explicitly and provide additional code there with the standard initialization
//code. You can evaluate the return value.
METHOD FB_Init: BOOL
VAR_INPUT
    bInitRetains: BOOL; // TRUE: the retain variables are initialized (reset warm / reset cold)
    bInCopyCode: BOOL;  // TRUE: the instance will be copied to the copy code afterward (online change)
    AxisRef    : REFERENCE TO AXIS_REF;
    iMotionStage : I_MotionStage;
END_VAR
THIS^.AxisRef REF= AxisRef;
THIS^.iMotionStage := iMotionStage ;
END_METHOD

METHOD Reset
VAR_INPUT
END_VAR
    fbTrigMgr.SetFrequency(fTargetFreq);
fbTrigMgr.ResetTriggerCounter();
nMoveIdx     := 0;
fSetpoint    := 0.0;
lastEndPoint := 0.0;
bStarted     := FALSE;
eState       := 0;
fbMoveAbs0.Execute := FALSE;
fbMoveAbs1.Execute := FALSE;
// Reset averaging state
bAvg    R= FALSE;
fSumPos := 0.0;
nSmpl   := 0;
fAvgPos := 0.0;
// Reset overshoot counters
nOvrCntPos := 0;
nOvrCntNeg := 0;
END_METHOD

METHOD Start
VAR_INPUT
END_VAR
fbTrigMgr.Stop();
fbMoveAbs0.Execute := FALSE;
fbMoveAbs1.Execute := FALSE;
IF ABS(iMotionStage.MotionStatus.fActPosition - fStopPos)
    < ABS(iMotionStage.MotionStatus.fActPosition - fStopNeg) THEN
    fSetpoint    := fStopPos;
    lastEndPoint := fStopPos;
ELSE
    fSetpoint    := fStopNeg;
    lastEndPoint := fStopNeg;
END_IF
fbTrigMgr.Start();
nMoveIdx := 0;
bStarted := TRUE;
END_METHOD

METHOD Stop
VAR_INPUT
END_VAR
fbTrigMgr.Stop();
fbMoveAbs0.Execute := FALSE;
fbMoveAbs1.Execute := FALSE;
eState   := 0;
bStarted := FALSE;
END_METHOD

END_FUNCTION_BLOCK

// ---- POUs/FB_TriggerManagerEL1124.TcPOU
FUNCTION_BLOCK FB_TriggerManagerEL1124 EXTENDS FB_TriggerManager
VAR
    bTriggerInputPrev       : BOOL := FALSE;
    nMinDebounceNs          : ULINT := 2000000; // 2 ms debounce in ns
    nLastTriggerTick        : ULINT := 0;
    nPrevTriggerTick        : ULINT := 0;
   {attribute 'pytmc' := '
        pv: fCurrentTriggerFrequency
        io: i
        field: DESC Current Trigger Frequency
    '}
    fCurrentTriggerFrequency : REAL := 0.0;
    nCurTick : ULINT := 0;
    nDeltaTick: ULINT;
END_VAR

IF (iTriggerSource = 0) THEN
    RETURN;
END_IF

nCurTick := F_GetCurDcTickTime64();

IF bRunning AND iTriggerSource.Trigger AND NOT bTriggerInputPrev THEN
    IF (nCurTick - nLastTriggerTick) >= nMinDebounceNs THEN
        bNewLatchPending := TRUE;
        nNumberOfTriggersSinceLastCounterReset := nNumberOfTriggersSinceLastCounterReset + 1;

        IF NOT bHaveNotReceivedFirstTriggerSinceLastStart THEN
            nDeltaTick := nCurTick - nPrevTriggerTick;
            IF nDeltaTick > 0 THEN
                fCurrentTriggerFrequency := 1.0 / (ULINT_TO_REAL(nDeltaTick) * 1E-9);
            ELSE
                fCurrentTriggerFrequency := fCurrentTriggerFrequency;
            END_IF
        ELSE
            bHaveNotReceivedFirstTriggerSinceLastStart := FALSE;
        END_IF

        nPrevTriggerTick := nCurTick;
        nLastTriggerTick := nCurTick;
    END_IF
END_IF

bTriggerInputPrev := iTriggerSource.Trigger;

END_FUNCTION_BLOCK

// ---- POUs/FB_MoveToNearestClosed.TcPOU
FUNCTION_BLOCK FB_MoveToNearestClosed
VAR_OUTPUT
    Closed   : BOOL;
END_VAR
VAR
    iMotionStage 		: I_MotionStage;
    fEndpointPositive  : LREAL :=  11.25;
    fEndpointNegative  : LREAL := -11.25;
    fTarget            : LREAL := 0.0;
    bStarted: BOOL;
END_VAR

Closed := FALSE;
IF 	bStarted THEN
    IF iMotionStage.MotionStatus.bDone THEN
        Closed := TRUE;
        bStarted := FALSE;
    END_IF
END_IF

//FB_Init is always available implicitly and it is used primarily for initialization.
//The return value is not evaluated. For a specific influence, you can also declare the
//methods explicitly and provide additional code there with the standard initialization
//code. You can evaluate the return value.
METHOD FB_Init: BOOL
VAR_INPUT
    bInitRetains: BOOL; // TRUE: the retain variables are initialized (reset warm / reset cold)
    bInCopyCode: BOOL;  // TRUE: the instance will be copied to the copy code afterward (online change)
    iMotionStage : I_MotionStage;
END_VAR
THIS^.iMotionStage := iMotionStage ;
END_METHOD

METHOD Start
// Choose closest endpoint
IF ABS(iMotionStage.MotionStatus.fActPosition - fEndpointPositive) < ABS(iMotionStage.MotionStatus.fActPosition - fEndpointNegative) THEN
    fTarget := fEndpointPositive;
ELSE
    fTarget := fEndpointNegative;
END_IF
// Issue move command
iMotionStage.AbsoluteMove(
   Position     := fTarget,
   Velocity     := iMotionStage.MotionCmd.fVelocity,
   Acceleration := iMotionStage.MotionCmd.fAcceleration,
   Deceleration := iMotionStage.MotionCmd.fDeceleration
);

bStarted := TRUE;
END_METHOD

END_FUNCTION_BLOCK

// ---- POUs/FB_FastOpen.TcPOU
FUNCTION_BLOCK  FB_FastOpen
VAR_INPUT
    fCenter	: LREAL;
END_VAR
VAR_OUTPUT
    Opened   : BOOL;
END_VAR

VAR
    iMotionStage	: I_MotionStage;
    bStarted : BOOL;
END_VAR

IF (iMotionStage = 0)  THEN
    RETURN;
END_IF

Opened := FALSE;
IF 	bStarted THEN
    IF iMotionStage.MotionStatus.bDone THEN
        Opened := TRUE;
        bStarted := FALSE;
    END_IF
END_IF

//FB_Init is always available implicitly and it is used primarily for initialization.
//The return value is not evaluated. For a specific influence, you can also declare the
//methods explicitly and provide additional code there with the standard initialization
//code. You can evaluate the return value.
METHOD FB_Init: BOOL
VAR_INPUT
    bInitRetains: BOOL; // TRUE: the retain variables are initialized (reset warm / reset cold)
    bInCopyCode: BOOL;  // TRUE: the instance will be copied to the copy code afterward (online change)
    iMotionStage : I_MotionStage;
END_VAR
THIS^.iMotionStage := iMotionStage ;
END_METHOD

METHOD Start : BOOL
VAR_INPUT
END_VAR
// Issue move command
iMotionStage.AbsoluteMoveDefault(
   Position     := fCenter,
   Velocity     := iMotionStage.MotionCmd.fVelocity,
);
bStarted := TRUE;
END_METHOD

END_FUNCTION_BLOCK

// ---- POUs/FB_FastClose.TcPOU
FUNCTION_BLOCK FB_FastClose
VAR_INPUT
    fStopPos : LREAL;
END_VAR
VAR_OUTPUT
    Closed   : BOOL;;
END_VAR
VAR
    iMotionStage       : I_MotionStage;
    bStarted : BOOL;
END_VAR

IF (iMotionStage = 0)  THEN
    RETURN;
END_IF

Closed := FALSE;
IF 	bStarted THEN
    IF iMotionStage.MotionStatus.bDone THEN
        Closed := TRUE;
        bStarted := FALSE;
    END_IF
END_IF

//FB_Init is always available implicitly and it is used primarily for initialization.
//The return value is not evaluated. For a specific influence, you can also declare the
//methods explicitly and provide additional code there with the standard initialization
//code. You can evaluate the return value.
METHOD FB_Init: BOOL
VAR_INPUT
    bInitRetains: BOOL; // TRUE: the retain variables are initialized (reset warm / reset cold)
    bInCopyCode: BOOL;  // TRUE: the instance will be copied to the copy code afterward (online change)
    iMotionStage : I_MotionStage;
END_VAR
THIS^.iMotionStage := iMotionStage ;
END_METHOD

METHOD Start : BOOL
VAR_INPUT
END_VAR
// Issue move command
iMotionStage.AbsoluteMoveDefault(
   Position     := fStopPos,
   Velocity     := iMotionStage.MotionCmd.fVelocity,
);
bStarted := TRUE;
END_METHOD

END_FUNCTION_BLOCK

// ---- POUs/FB_SpindleHomeToCenter.TcPOU
(*  FB_HomeIndex - Index pulse homing sequence for the spindle.

 Overview:
   Manages a multi-state homing sequence that uses a physical index pulse
   (bHomeIndex) to establish a reference position. On detecting a homing
   start, the FB waits for the index pulse, latches a HomeLimit signal for
   a configurable duration, then waits for the drive to confirm homed+done
   before issuing a centering move to fCenterOffset. Finally it zeros the
   position via MC_SetPosition and enables backlash compensation.
*)
FUNCTION_BLOCK FB_SpindleHomeToCenter
VAR_INPUT
    fCenterOffset : LREAL;
    fDefaultVelocity : LREAL;
END_VAR
VAR
    iMotionStage 		: I_MotionStage;
    bHomeIndex  AT %I* : BOOL;
    {attribute 'hide'}
    rtHomingStart     : R_TRIG;
    {attribute 'hide'}
    rtHomePulse       : R_TRIG;
    {attribute 'hide'}
    rtDoneHome        : R_TRIG;
    {attribute 'hide'}
    rtCenterDone       : R_TRIG;
    {attribute 'hide'}
    rtError : R_TRIG;

    nCurTick          : ULINT;
    nLatchStartTick   : ULINT;
    nLatchDurationNs  : ULINT := 30_000_000; // 30ms (adjust as needed)
    bHomePulseLatched : BOOL;
    fPrevVelocity     : LREAL;
    fbMcSetPosition   : MC_SetPosition;


    rtHomed: R_TRIG;
    rtWaitHomeIndexDone: R_TRIG;
END_VAR

VAR_OUTPUT
   {attribute 'pytmc' := '
        pv: bCentered
        io: i
        field: ZNAM FALSE
        field: ONAM TRUE
        field: DESC TRUE if the pulse picker is centered
    '}
    bCentered   : BOOL;
    bHomeDone         : BOOL;
    bLocalError       : BOOL;
    eHomeIndexState : E_HomeIndexState := E_HomeIndexState.Idle;
END_VAR

IF (iMotionStage = 0) THEN
    RETURN;
END_IF

nCurTick := F_GetCurDcTickTime64();

rtError(CLK := iMotionStage.MotionStatus.bError AND iMotionStage.MotionStatus.bStageReady);
rtHomingStart(CLK := iMotionStage.MotionStatus.bHoming);
rtHomePulse(CLK := bHomeIndex);
rtHomed(CLK := iMotionStage.MotionStatus.bHomed);
// Fires when drive confirms both done and homed after index pulse
rtWaitHomeIndexDone(CLK := iMotionStage.MotionStatus.bDone
        AND iMotionStage.MotionStatus.bHomed
        AND (eHomeIndexState = E_HomeIndexState.WaitHomeDone));
// Fires when centering alignment move completes
rtCenterDone(CLK := iMotionStage.MotionStatus.bDone
    AND (eHomeIndexState = E_HomeIndexState.CenterMove));

// Any drive error immediately redirects to Error state from any point in sequence
IF rtError.Q THEN
    eHomeIndexState := E_HomeIndexState.Error;
END_IF

